{region 'Documentation'}
(*!
<summary>Evaluates captured observations after the scenario has finished.</summary>
*)
{endregion}
METHOD PROTECTED ProcessAssertions
VAR_INPUT
    Enable : BOOL; //! Phase permission supplied by the owning Test Case; FALSE does not authorize progression, while observation may continue.
END_VAR
VAR
    Evaluate : BOOL;
END_VAR
Evaluate := Enable AND FPerformed;
FActiveRun(Enable := Evaluate,
    State := State,
    IN := FActiveRunMatches);
FResetBoundary(Enable := Evaluate,
    State := State,
    IN := FResetBoundaryMatches);
FReservationsReleased(Enable := Evaluate,
    State := State,
    IN := FReservationsReleasedMatches);
FErrorPath(Enable := Evaluate,
    State := State,
    IN := FErrorPathMatches);
FNoLifecycleReset(Enable := Evaluate,
    State := State,
    IN := FNoLifecycleResetMatches);
FNewEpoch(Enable := Evaluate,
    State := State,
    IN := FNewEpochMatches);
FFinalization(Enable := Evaluate,
    State := State,
    IN := FFinalizationMatches);
FConfigurationPreserved(Enable := Evaluate,
    State := State,
    IN := FConfigurationPreservedMatches);
IF Evaluate THEN
    FChecked := TRUE;
END_IF;
END_METHOD

{region 'Documentation'}
(*!
<summary>No Preparation phase is needed.</summary>
*)
{endregion}
METHOD PROTECTED ProcessPreparations
VAR_INPUT
    // SA0033: Required override without Preparation work.
    {attribute 'analysis' := '-33'}
    Enable : BOOL; //! Phase permission supplied by the owning Test Case; FALSE does not authorize progression, while observation may continue.
END_VAR
END_METHOD

{region 'Documentation'}
(*!
<summary>Resets observations and schedules a fresh subject initialization.</summary>
*)
{endregion}
METHOD PROTECTED ProcessReset
FPerformed := FALSE;
FChecked := FALSE;
FPhase := SetupPhase;
FSuite := 0;
FChild := 0;
FSecondChild := 0;
FActiveRun.Reset();
FActiveRunMatches := FALSE;
FResetBoundary.Reset();
FResetBoundaryMatches := FALSE;
FReservationsReleased.Reset();
FReservationsReleasedMatches := FALSE;
FErrorPath.Reset();
FErrorPathMatches := FALSE;
FNoLifecycleReset.Reset();
FNoLifecycleResetMatches := FALSE;
FNewEpoch.Reset();
FNewEpochMatches := FALSE;
FFinalization.Reset();
FFinalizationMatches := FALSE;
FConfigurationPreserved.Reset();
FConfigurationPreservedMatches := FALSE;
CompleteReset();
END_METHOD

{region 'Documentation'}
(*!
<summary>Runs the bounded scenario once before Assertion evaluation.</summary>
*)
{endregion}
METHOD PROTECTED ProcessTests
VAR_INPUT
    Enable : BOOL; //! Phase permission supplied by the owning Test Case; FALSE does not authorize progression, while observation may continue.
END_VAR
IF NOT Enable THEN
    RETURN;
END_IF;
IF FChecked THEN
    CompleteTests();
    RETURN;
END_IF;

IF NOT FPerformed THEN
    StateMachine();
END_IF;
END_METHOD

{region 'Documentation'}
(*!
<summary>Advances the real hierarchy once per cycle and separates reset boundary from error completion.</summary>
*)
{endregion}
METHOD PRIVATE StateMachine
VAR
    EmptyControl : ST_RunControl;
    SeedEvent : ST_Event;
    Published : INT;
END_VAR
CASE FPhase OF
    SetupPhase:
        FControl := EmptyControl;
        IF NOT FSubject.Initialize(Buffer := FEvents,
            FifoControl := FFifo,
            Status := FBufferStatus) THEN
            Error(Message := 'Active reset buffer initialization failed.');
            RETURN;
        END_IF;
        FRoot.BindPublisher(Publisher := FSubject);
        IF NOT FRoot.Initialize(Name := 'ActiveReset',
            EventBuffer := FSubject) THEN
            Error(Message := 'Active reset hierarchy initialization failed.');
            RETURN;
        END_IF;
        FSuite := FRoot.GetTestSuite(Index := FRoot.ChildArrayLowerBound);
        FChild := FRoot.GetTestCase(Index := FRoot.TestCaseLowerBound);
        FSecondChild := FRoot.GetTestCase(Index := FRoot.TestCaseLowerBound + 1);
        IF (FSuite = 0) OR (FChild = 0) OR (FSecondChild = 0) THEN
            Error(Message := 'Active reset hierarchy is incomplete.');
            RETURN;
        END_IF;
        FPhase := AwaitIdlePhase;

    AwaitIdlePhase:
        FRoot(ControlData := FControl);
        IF FRoot.HasError THEN
            Error(Message := 'Active reset hierarchy did not establish Idle.');
            RETURN;
        END_IF;
        IF FRoot.IsReady THEN
            FRoot.RequestStart();
            FPhase := AwaitActivePhase;
        END_IF;

    AwaitActivePhase:
        FRoot(ControlData := FControl);
        IF FRoot.HasError OR FRoot.IsComplete THEN
            Error(Message := 'Hierarchy ended before the active reset precondition.');
            RETURN;
        END_IF;
        IF FChild.State = E_State.Running THEN
            FActiveRunMatches := (FRoot.State = E_State.Running) AND (FSuite.State = E_State.Running)
                AND (FSuite.ReservedEntryCount > 0) AND (FChild.ReservedEntryCount > 0)
                AND (FSubject.ReservedEntryCount > 0);
            SeedEvent := CreateFrameworkEvent(Name := 'ActiveReset',
                ResourceName := 'ActiveResetFixture',
                State := E_State.Running,
                Severity := E_EventSeverity.Info,
                Message := OldEpochMarker);
            Published := FSubject.PublishEvent(Event := SeedEvent);
            FActiveRunMatches := FActiveRunMatches AND (Published > 0);
            FSubject.Arm(Root := FRoot,
                Suite := FSuite,
                Child := FChild);
            FPhase := ResetPhase;
        END_IF;

    ResetPhase:
        FControl.BufferCmd.Reset := TRUE;
        FRoot(ControlData := FControl);
        FResetBoundaryMatches := FSubject.Observed AND FSubject.LifecycleUnchanged
            AND FSubject.EpochCleared AND NOT FControl.BufferCmd.Reset
            AND (FControl.BufferCmd.DeleteSequenceId = 0);
        FReservationsReleasedMatches := FSubject.OwnersReleased
            AND (FSuite.ReservedEntryCount = 0) AND (FChild.ReservedEntryCount = 0)
            AND (FSecondChild.ReservedEntryCount = 0);
        FPhase := AwaitCompletionPhase;

    AwaitCompletionPhase:
        FRoot(ControlData := FControl);
        IF FRoot.IsComplete THEN
            CheckNewEpoch();
            FFinalizationMatches := FFinalizationMatches AND (FRoot.Result = E_Result.Error)
                AND FRoot.HasError;
            FConfigurationPreservedMatches := FRoot.ConfigurationUnchanged AND FRoot.ChildCallsMatch;
            FPerformed := TRUE;
        END_IF;

    ELSE
        Error(Message := 'Unknown active buffer reset phase.');
END_CASE;
END_METHOD

END_FUNCTION_BLOCK

// ---- SelfTests/TestCases/TestSuite_EventBufferReset/Helper/ActiveResetBufferProbe.TcPOU
{region 'Documentation'}
(*!
<summary>Records the synchronous hard-reset boundary before the owner resumes lifecycle processing.</summary>
<description>
Arm captures the real active hierarchy. Reset delegates storage handling unchanged to EventBuffer,
then records cleared metadata and unchanged lifecycle states. Subsequent owner processing may
legitimately publish errors and request Abort; those actions are outside this observation boundary.
Initialization resets are ignored until Arm. The test keeps all referenced objects alive.
</description>
*)
{endregion}
FUNCTION_BLOCK ActiveResetBufferProbe EXTENDS EventBuffer
VAR
    FArmed : BOOL;
    FRoot : REFERENCE TO RunControlIntegrationSubject;
    FSuite : I_TestSuite;
    FChild : I_TestCase;
    FRootState : E_State;
    FSuiteState : E_State;
    FChildState : E_State;
    FLifecycleUnchanged : BOOL;
    FEpochCleared : BOOL;
    FOwnersReleased : BOOL;
    FObserved : BOOL;
END_VAR

{region 'Documentation'}
(*!
<summary>Captures the active hierarchy immediately before the external Buffer Reset.</summary>
*)
{endregion}
METHOD PUBLIC Arm
VAR_INPUT
    Suite : I_TestSuite; //! Borrowed Suite observed across the Reset boundary; keep it alive while armed.
    Child : I_TestCase; //! Borrowed child observed across the Reset boundary; keep it alive while armed.
END_VAR
VAR_IN_OUT
    // SA0167: Borrowed real owner, retained only for state observations.
    {attribute 'analysis' := '-167'}
    Root : RunControlIntegrationSubject; //! Borrowed real Run-Control owner retained for state observations; keep it alive while armed.
END_VAR
FRoot REF= Root;
FSuite := Suite;
FChild := Child;
FRootState := Root.State;
FSuiteState := Suite.State;
FChildState := Child.State;
FLifecycleUnchanged := FALSE;
FEpochCleared := FALSE;
FOwnersReleased := FALSE;
FObserved := FALSE;
FArmed := TRUE;
END_METHOD

{region 'Documentation'}
(*!
<summary>Recorded EpochCleared for command-order verification.</summary>
*)
{endregion}
{attribute 'monitoring' := 'call'}
PROPERTY PUBLIC EpochCleared : BOOL //! Recorded EpochCleared for command-order verification.
GET
EpochCleared := FEpochCleared;
END_GET
END_PROPERTY

{region 'Documentation'}
(*!
<summary>Recorded LifecycleUnchanged for command-order verification.</summary>
*)
{endregion}
{attribute 'monitoring' := 'call'}
PROPERTY PUBLIC LifecycleUnchanged : BOOL //! Recorded LifecycleUnchanged for command-order verification.
GET
LifecycleUnchanged := FLifecycleUnchanged;
END_GET
END_PROPERTY

{region 'Documentation'}
(*!
<summary>Recorded Observed for command-order verification.</summary>
*)
{endregion}
{attribute 'monitoring' := 'call'}
PROPERTY PUBLIC Observed : BOOL //! Recorded Observed for command-order verification.
GET
Observed := FObserved;
END_GET
END_PROPERTY

{region 'Documentation'}
(*!
<summary>Recorded OwnersReleased for command-order verification.</summary>
*)
{endregion}
{attribute 'monitoring' := 'call'}
PROPERTY PUBLIC OwnersReleased : BOOL //! Recorded OwnersReleased for command-order verification.
GET
OwnersReleased := FOwnersReleased;
END_GET
END_PROPERTY

{region 'Documentation'}
(*!
<summary>Delegates real reset and snapshots its immediate effects, not later owner processing.</summary>
*)
{endregion}
METHOD PUBLIC Reset
VAR
    Epoch : ST_EventBufferStatus;
    CurrentFifoStatus : ST_FifoStatus;
END_VAR
IF FArmed THEN
    FOwnersReleased := (FSuite.ReservedEntryCount = 0) AND (FChild.ReservedEntryCount = 0)
        AND (ReservedEntryCount = 0);
END_IF;
SUPER^.Reset();
IF FArmed THEN
    Epoch := Status;
    CurrentFifoStatus := FifoStatus;
    FEpochCleared := CurrentFifoStatus.BufferEmpty AND (CurrentFifoStatus.ElementCount = 0)
        AND (Epoch.SequenceId = 0) AND (Epoch.DeletedSequenceId = 0)
        AND (Epoch.LostEventCount = 0) AND (ReservedEntryCount = 0);
    FLifecycleUnchanged := (FRoot.State = FRootState) AND (FSuite.State = FSuiteState)
        AND (FChild.State = FChildState);
    FObserved := TRUE;
    FArmed := FALSE;
END_IF;
END_METHOD

END_FUNCTION_BLOCK

// ---- SelfTests/TestSuites/TestSuite_AssertionLifecycle.TcPOU
{region 'Documentation'}
(*!
<summary>Checks shared Assertion identity, activity, reset and result-event behavior.</summary>
*)
{endregion}
FUNCTION_BLOCK TestSuite_AssertionLifecycle EXTENDS TestSuiteBase
VAR
    FInitialization : Test_AssertionInitialization;
    FActivity : Test_AssertionActivity;
    FUninitialized : Test_AssertionUninitialized;
    FResetReuse : Test_AssertionResetReuse;
    FEscalation : Test_AssertionEscalation;
    FTestCases : ARRAY[1..TestCaseCapacity] OF I_TestCase;
END_VAR
VAR CONSTANT
    TestCaseCapacity : UINT := 5;
END_VAR

SUPER^();

{region 'Documentation'}
(*!
<summary>Initializes and registers the five isolated Assertion lifecycle scenarios.</summary>
*)
{endregion}
METHOD PROTECTED Configure
VAR_IN_OUT
    // SA0167: Borrowed owner builder; no temporary instance is created.
    {attribute 'analysis' := '-167'}
    Builder : TestSuiteConfigurationBuilder; //! Borrowed owner configuration builder used only during this Configure call; register this owner's concrete children.
END_VAR
VAR
    TestConfig : ST_TestCaseConfig;
END_VAR
Builder.Initialize(Mode := E_OrchestrationMode.Serial,
    TestCases := FTestCases);
FInitialization.Initialize(Parent := THIS^,
    TestName := 'Initialization',
    Config := TestConfig);
Builder.Register(TestCase := FInitialization);
FActivity.Initialize(Parent := THIS^,
    TestName := 'Activity',
    Config := TestConfig);
Builder.Register(TestCase := FActivity);
FUninitialized.Initialize(Parent := THIS^,
    TestName := 'Uninitialized',
    Config := TestConfig);
Builder.Register(TestCase := FUninitialized);
FResetReuse.Initialize(Parent := THIS^,
    TestName := 'ResetReuse',
    Config := TestConfig);
Builder.Register(TestCase := FResetReuse);
FEscalation.Initialize(Parent := THIS^,
    TestName := 'Escalation',
    Config := TestConfig);
Builder.Register(TestCase := FEscalation);
END_METHOD

{region 'Documentation'}
(*!
<summary>Returns a registered scenario using its original array index.</summary>
*)
{endregion}
METHOD PUBLIC GetTestCase : I_TestCase //! Typed child interface at the original array index; zero when no entry is available.
VAR_INPUT
    Index : DINT; //! Original occupied child-array index, rather than an ordinal position.
END_VAR
GetTestCase := 0;
IF (ChildCount = 0) OR (Index < ChildArrayLowerBound)
    OR (DINT_TO_LINT(Index) >= DINT_TO_LINT(ChildArrayLowerBound) + UINT_TO_LINT(ChildCount)) THEN
    RETURN;
END_IF;
GetTestCase := FTestCases[Index];
END_METHOD

{region 'Documentation'}
(*!
<summary>Calls each owned scenario once per initialized Suite cycle.</summary>
*)
{endregion}
METHOD PROTECTED ProcessTestCases
FInitialization();
FActivity();
FUninitialized();
FResetReuse();
FEscalation();
END_METHOD

END_FUNCTION_BLOCK

// ---- SelfTests/TestCases/TestSuite_AssertionLifecycle/Test_AssertionInitialization.TcPOU
{region 'Documentation'}
(*!
<summary>Checks Assertion identity validation and deferred reset dispatch.</summary>
<description>
Each attempt changes one identity/configuration condition. Initialize is checked before
any FB call; three later calls verify reset dispatch, valid activity or rejected passivity.
Checking Assertions latch every attempt, while intentional diagnostics stay local.
Publisher checks cover zero rejection, explicit replacement and unchanged lifecycle/history
before and after subject calls. A separate untouched Assertion verifies the lazy default.
Repeated runs use the same subject and reinitialize it; they do not claim fresh memory.
</description>
*)
{endregion}
FUNCTION_BLOCK Test_AssertionInitialization EXTENDS TestCaseBase
VAR
    FSubject : AssertionLifecycleSubject;
    FDefaultSubject : AssertTrue;
    FAlternativeCapture : EventBuffer;
    FAlternativeEvents : ARRAY[1..CaptureLength] OF ST_Event;
    FAlternativeFifo : ST_FifoStatus;
    FAlternativeStatus : ST_EventBufferStatus;
    FParent : AssertionParentIdentity;
    FCapture : EventBuffer;
    FEvents : ARRAY[1..CaptureLength] OF ST_Event;
    FCaptureFifo : ST_FifoStatus;
    FCaptureStatus : ST_EventBufferStatus;
    FAttempt : UINT;
    FCall : UINT;
    FAttemptStarted : BOOL;
    FExpectedInitialized : BOOL;
    FExpectedObserveFirstCycle : BOOL;
    FExpectedName : STRING(GVL_Constants.NameLength);
    FExpectedResource : STRING(GVL_Constants.ResourceNameLength);
    FExpectedEvents : UDINT;
    FObservationReady : BOOL;
    FChecked : BOOL;
END_VAR
VAR
    FPublisherBinding : AssertTrue;
    FPublisherBindingMatches : BOOL;
    FInitialization : AssertTrue;
    FInitializationMatches : BOOL;
    FIdentity : AssertTrue;
    FIdentityMatches : BOOL;
    FSettings : AssertTrue;
    FSettingsMatches : BOOL;
    FDispatch : AssertTrue;
    FDispatchMatches : BOOL;
    FActivity : AssertTrue;
    FActivityMatches : BOOL;
    FDiagnostics : AssertTrue;
    FDiagnosticsMatches : BOOL;
    FCaptureIntegrity : AssertTrue;
    FCaptureIntegrityMatches : BOOL;
END_VAR
VAR CONSTANT
    CaptureLength : UINT := 8;
    DefaultSettings : UINT := 1;
    DottedSuffix : UINT := 2;
    ExactCapacity : UINT := 3;
    OverCapacity : UINT := 4;
    MissingParent : UINT := 5;
    EmptySuffix : UINT := 6;
    InvalidParent : UINT := 7;
    NonAsciiSuffix : UINT := 8;
    ExplicitSettings : UINT := 9;
    LastAttempt : UINT := ExplicitSettings;
    ResetCall : UINT := 1;
    SecondCheckCall : UINT := 3;
    ResetSampleValue : UINT := 17;
END_VAR

SUPER^();

{region 'Documentation'}
(*!
<summary>Collects only outer checking Assertions, never intentional subject findings.</summary>
*)
{endregion}
METHOD PROTECTED AggregateResults
VAR_INPUT
    Aggregator : I_ResultAggregator; //! Borrowed result sink owned by the outer Test Case; add this test's checking Assertions without resetting or retaining the sink.
END_VAR
Aggregator.AddProvider(Provider := FPublisherBinding);
Aggregator.AddProvider(Provider := FInitialization);
Aggregator.AddProvider(Provider := FIdentity);
Aggregator.AddProvider(Provider := FSettings);
Aggregator.AddProvider(Provider := FDispatch);
Aggregator.AddProvider(Provider := FActivity);
Aggregator.AddProvider(Provider := FDiagnostics);
Aggregator.AddProvider(Provider := FCaptureIntegrity);
END_METHOD

{region 'Documentation'}
(*!
<summary>Varies one setup condition and observes Initialize before cyclic processing.</summary>
*)
{endregion}
METHOD PRIVATE BeginAttempt
VAR
    Parent : I_TestCase;
    ParentName : STRING(GVL_Constants.NameLength);
    LocalName : STRING(GVL_Constants.NameLength);
    FullName : STRING(2 * GVL_Constants.NameLength + 1);
    Initialized : BOOL;
    SuffixLength : INT;
    Index : INT;
END_VAR
IF NOT FCapture.Initialize(Buffer := FEvents,
    FifoControl := FCaptureFifo,
    Status := FCaptureStatus) THEN
    Error(Message := 'Assertion initialization capture setup failed.');
    RETURN;
END_IF;

IF NOT FAlternativeCapture.Initialize(Buffer := FAlternativeEvents,
    FifoControl := FAlternativeFifo,
    Status := FAlternativeStatus) THEN
    Error(Message := 'Alternative Assertion publisher setup failed.');
    RETURN;
END_IF;

CheckPublisherBinding();
ParentName := 'Root.Suite.Case';
LocalName := 'Subject';
FExpectedInitialized := TRUE;
FExpectedObserveFirstCycle := TRUE;
FExpectedResource := '';
CASE FAttempt OF
    DefaultSettings:
        LocalName := 'Subject';
    DottedSuffix:
        LocalName := 'Value.With.Detail';
    ExactCapacity, OverCapacity:
        LocalName := '';
        SuffixLength := UINT_TO_INT(GVL_Constants.NameLength) - LEN(ParentName) - 1;
        IF FAttempt = OverCapacity THEN
            SuffixLength := SuffixLength + 1;
            FExpectedInitialized := FALSE;
        END_IF;
        FOR Index := 1 TO SuffixLength DO
            LocalName := CONCAT(LocalName, 'x');
        END_FOR;
    MissingParent:
        FExpectedInitialized := FALSE;
    EmptySuffix:
        LocalName := '';
        FExpectedInitialized := FALSE;
    InvalidParent:
        ParentName := 'Root..Case';
        FExpectedInitialized := FALSE;
    NonAsciiSuffix:
        // SA0175: Deliberately invalid non-ASCII identity input for the rejection test.
        {analysis -175}
        LocalName := '$E4';
        {analysis +175}
        FExpectedInitialized := FALSE;
    ExplicitSettings:
        FExpectedResource := 'Resource';
        FExpectedObserveFirstCycle := FALSE;
ELSE
    Error(Message := 'Unknown Assertion initialization attempt.');
    RETURN;
END_CASE;

FParent.SetIdentity(Value := ParentName);
Parent := FParent;
IF FAttempt = MissingParent THEN
    Parent := 0;
    FExpectedName := LocalName;
ELSE
    FullName := CONCAT(CONCAT(ParentName, '.'), LocalName);
    // SA0175: The expected diagnostic projection is deliberately bounded ASCII-byte truncation.
    {analysis -175}
    FExpectedName := LEFT(FullName, UINT_TO_INT(GVL_Constants.NameLength));
    {analysis +175}
END_IF;

FSubject.ClearTrace();
IF FAttempt = ExplicitSettings THEN
    Initialized := FSubject.Initialize(Parent := Parent,
        AssertionName := LocalName,
        ResourceName := FExpectedResource,
        ObserveFirstCycle := FExpectedObserveFirstCycle);
ELSE
    Initialized := FSubject.Initialize(Parent := Parent,
        AssertionName := LocalName);
END_IF;
FInitializationMatches := (Initialized = FExpectedInitialized)
    AND (FSubject.IsInitialized = FExpectedInitialized)
    AND (FSubject.Result = E_Result.NotEvaluated);
FIdentityMatches := TRUE;
FSettingsMatches := TRUE;
IF FAttempt <> MissingParent THEN
    FIdentityMatches := FSubject.Name = FExpectedName;
    FSettingsMatches := (FSubject.ResourceName = FExpectedResource)
        AND (FSubject.ObserveFirstCycle = FExpectedObserveFirstCycle);
END_IF;
FDispatchMatches := (FSubject.ResetCallCount = 0) AND (FSubject.AssertCallCount = 0);
FActivityMatches := NOT FSubject.Enabled
    AND NOT FSubject.ObservationActive AND NOT FSubject.EvaluationActive;
FExpectedEvents := 0;
FDiagnosticsMatches := TRUE;
IF NOT FExpectedInitialized THEN
    FExpectedEvents := 1;
    FDiagnosticsMatches := (FEvents[1].Name = FExpectedName)
        AND (FEvents[1].OwnerScope = E_OwnerScope.Framework)
        AND (FEvents[1].EventType = E_EventType.Framework)
        AND (FEvents[1].Severity = E_EventSeverity.Error)
        AND (FEvents[1].State = E_State.Uninitialized);
END_IF;
FDiagnosticsMatches := FDiagnosticsMatches AND (FCaptureStatus.SequenceId = FExpectedEvents);
FCaptureIntegrityMatches := FCaptureStatus.LostEventCount = 0;
FAttemptStarted := TRUE;
FCall := ResetCall;
END_METHOD

{region 'Documentation'}
(*!
<summary>Checks binding without changing subject lifecycle, history or event counts.</summary>
*)
{endregion}
METHOD PRIVATE CheckPublisherBinding
VAR
    PrimaryPublisher : I_EventPublisher;
    AlternativePublisher : I_EventPublisher;
    DefaultPublisher : I_EventPublisher;
    ResultBefore : E_Result;
    InitializedBefore : BOOL;
    EnabledBefore : BOOL;
    ObservationBefore : BOOL;
    EvaluationBefore : BOOL;
    NameBefore : STRING(GVL_Constants.NameLength);
    SequenceBefore : UDINT;
    AlternativeSequenceBefore : UDINT;
END_VAR
PrimaryPublisher := FCapture;
AlternativePublisher := FAlternativeCapture;
DefaultPublisher := GVL_EventBuffer.Publisher;
FDefaultSubject.BindPublisher(Publisher := 0);
FPublisherBindingMatches := FPublisherBindingMatches
    AND (FDefaultSubject.EventPublisher = DefaultPublisher);

ResultBefore := FSubject.Result;
InitializedBefore := FSubject.IsInitialized;
EnabledBefore := FSubject.Enabled;
ObservationBefore := FSubject.ObservationActive;
EvaluationBefore := FSubject.EvaluationActive;
NameBefore := FSubject.Name;
SequenceBefore := FCaptureStatus.SequenceId;
AlternativeSequenceBefore := FAlternativeStatus.SequenceId;

FSubject.BindPublisher(Publisher := AlternativePublisher);
FPublisherBindingMatches := FPublisherBindingMatches
    AND (FSubject.EventPublisher = AlternativePublisher);
FSubject.BindPublisher(Publisher := 0);
FPublisherBindingMatches := FPublisherBindingMatches
    AND (FSubject.EventPublisher = AlternativePublisher);
FSubject.BindPublisher(Publisher := PrimaryPublisher);
FPublisherBindingMatches := FPublisherBindingMatches
    AND (FSubject.EventPublisher = PrimaryPublisher)
    AND (FSubject.Result = ResultBefore)
    AND (FSubject.IsInitialized = InitializedBefore)
    AND (FSubject.Enabled = EnabledBefore)
    AND (FSubject.ObservationActive = ObservationBefore)
    AND (FSubject.EvaluationActive = EvaluationBefore)
    AND (FSubject.Name = NameBefore)
    AND (FCaptureStatus.SequenceId = SequenceBefore)
    AND (FAlternativeStatus.SequenceId = AlternativeSequenceBefore);
END_METHOD

{region 'Documentation'}
(*!
<summary>Configures checking Assertions; subject actions remain in the test script.</summary>
*)
{endregion}
METHOD PROTECTED Configure
FPreparationStateCount := 0;
FTestStateCount := 1;
FPublisherBinding.Initialize(Parent := THIS^,
    AssertionName := 'PublisherBinding');
FInitialization.Initialize(Parent := THIS^,
    AssertionName := 'Initialization');
FIdentity.Initialize(Parent := THIS^,
    AssertionName := 'Identity');
FSettings.Initialize(Parent := THIS^,
    AssertionName := 'Settings');
FDispatch.Initialize(Parent := THIS^,
    AssertionName := 'Dispatch');
FActivity.Initialize(Parent := THIS^,
    AssertionName := 'Activity');
FDiagnostics.Initialize(Parent := THIS^,
    AssertionName := 'Diagnostics');
FCaptureIntegrity.Initialize(Parent := THIS^,
    AssertionName := 'CaptureIntegrity');
FSubject.BindPublisher(Publisher := FCapture);
END_METHOD

{region 'Documentation'}
(*!
<summary>Checks reset and subsequent dispatch using one subject call per cycle.</summary>
*)
{endregion}
METHOD PRIVATE ObserveCall
VAR
    ExpectedActive : BOOL;
END_VAR
FSubject(Enable := TRUE,
    State := E_State.Running,
    Sample := ResetSampleValue);
FDispatchMatches := FDispatchMatches
    AND (FSubject.ResetCallCount = 1) AND (FSubject.ResetSample = ResetSampleValue);
IF FCall = ResetCall THEN
    FDispatchMatches := FDispatchMatches AND (FSubject.AssertCallCount = 0)
        AND (FSubject.ObservedSample = 0);
    FActivityMatches := FActivityMatches AND FSubject.Enabled
        AND NOT FSubject.ObservationActive AND NOT FSubject.EvaluationActive
        AND (FSubject.Result = E_Result.NotEvaluated);
ELSIF FExpectedInitialized THEN
    FDispatchMatches := FDispatchMatches AND (FSubject.AssertCallCount = FCall - 1);
    ExpectedActive := FExpectedObserveFirstCycle OR (FCall = SecondCheckCall);
    FActivityMatches := FActivityMatches AND FSubject.Enabled
        AND (FSubject.ObservationActive = ExpectedActive)
        AND (FSubject.EvaluationActive = ExpectedActive);
    IF ExpectedActive THEN
        FActivityMatches := FActivityMatches AND (FSubject.Result = E_Result.Passed);
    ELSE
        FActivityMatches := FActivityMatches AND (FSubject.Result = E_Result.NotEvaluated);
    END_IF;
ELSE
    FDispatchMatches := FDispatchMatches AND (FSubject.AssertCallCount = 0);
    FActivityMatches := FActivityMatches AND NOT FSubject.ObservationActive
        AND NOT FSubject.EvaluationActive AND (FSubject.Result = E_Result.NotEvaluated);
END_IF;
FDiagnosticsMatches := FDiagnosticsMatches AND (FCaptureStatus.SequenceId = FExpectedEvents);
FCaptureIntegrityMatches := FCaptureIntegrityMatches AND (FCaptureStatus.LostEventCount = 0);
CheckPublisherBinding();
FObservationReady := TRUE;
END_METHOD

{region 'Documentation'}
(*!
<summary>Completes abort without asynchronous resources.</summary>
*)
{endregion}
METHOD PROTECTED ProcessAbort
VAR_INPUT
    Enable : BOOL; //! Phase permission supplied by the owning Test Case; FALSE does not authorize progression, while observation may continue.
END_VAR
IF Enable THEN
    CompleteAbort();
END_IF;
END_METHOD

{region 'Documentation'}
(*!
<summary>Latches checked observations before the next script step may proceed.</summary>
*)
{endregion}
METHOD PROTECTED ProcessAssertions
VAR_INPUT
    Enable : BOOL; //! Phase permission supplied by the owning Test Case; FALSE does not authorize progression, while observation may continue.
END_VAR
VAR
    Evaluate : BOOL;
END_VAR
Evaluate := Enable AND FObservationReady;
FPublisherBinding(Enable := Evaluate,
    State := State,
    IN := FPublisherBindingMatches);
FInitialization(Enable := Evaluate,
    State := State,
    IN := FInitializationMatches);
FIdentity(Enable := Evaluate,
    State := State,
    IN := FIdentityMatches);
FSettings(Enable := Evaluate,
    State := State,
    IN := FSettingsMatches);
FDispatch(Enable := Evaluate,
    State := State,
    IN := FDispatchMatches);
FActivity(Enable := Evaluate,
    State := State,
    IN := FActivityMatches);
FDiagnostics(Enable := Evaluate,
    State := State,
    IN := FDiagnosticsMatches);
FCaptureIntegrity(Enable := Evaluate,
    State := State,
    IN := FCaptureIntegrityMatches);
IF Evaluate THEN
    FChecked := TRUE;
END_IF;
END_METHOD

{region 'Documentation'}
(*!
<summary>No Preparation phase is required.</summary>
*)
{endregion}
METHOD PROTECTED ProcessPreparations
VAR_INPUT
    // SA0033: Required hook; this test has no Preparation phase.
    {attribute 'analysis' := '-33'}
    Enable : BOOL; //! Phase permission supplied by the owning Test Case; FALSE does not authorize progression, while observation may continue.
END_VAR
END_METHOD

{region 'Documentation'}
(*!
<summary>Restarts the script and resets the checking Assertions.</summary>
*)
{endregion}
METHOD PROTECTED ProcessReset
FPublisherBinding.Reset();
FPublisherBindingMatches := TRUE;
FAttempt := DefaultSettings;
FCall := ResetCall;
FAttemptStarted := FALSE;
FObservationReady := FALSE;
FChecked := FALSE;
FInitialization.Reset();
FInitializationMatches := TRUE;
FIdentity.Reset();
FIdentityMatches := TRUE;
FSettings.Reset();
FSettingsMatches := TRUE;
FDispatch.Reset();
FDispatchMatches := TRUE;
FActivity.Reset();
FActivityMatches := TRUE;
FDiagnostics.Reset();
FDiagnosticsMatches := TRUE;
FCaptureIntegrity.Reset();
FCaptureIntegrityMatches := TRUE;
CompleteReset();
END_METHOD

{region 'Documentation'}
(*!
<summary>Advances one bounded script step per active PLC cycle.</summary>
*)
{endregion}
METHOD PROTECTED ProcessTests
VAR_INPUT
    Enable : BOOL; //! Phase permission supplied by the owning Test Case; FALSE does not authorize progression, while observation may continue.
END_VAR
IF NOT Enable THEN
    RETURN;
END_IF;
IF FChecked THEN
    FChecked := FALSE;
    FObservationReady := FALSE;
    IF FCall = SecondCheckCall THEN
        IF FAttempt = LastAttempt THEN
            CompleteTests();
            RETURN;
        END_IF;
        FAttempt := FAttempt + 1;
        FAttemptStarted := FALSE;
    ELSE
        FCall := FCall + 1;
    END_IF;
END_IF;
IF NOT FAttemptStarted THEN
    BeginAttempt();
    RETURN;
END_IF;
ObserveCall();
END_METHOD

END_FUNCTION_BLOCK

// ---- SelfTests/TestCases/TestSuite_AssertionLifecycle/Helper/AssertionLifecycleSubject.TcPOU
{region 'Documentation'}
(*!
<summary>Exposes calls and activity gates of AssertionBase without replacing its processing.</summary>
<description>
Bind the local publisher before Initialize. The inherited body owns initialization,
reset priority and activity history. Assert records both gates and a bounded sample;
active evaluation dispatches the selected inherited finding method without a result guard.
This deliberately exercises base-owned suppression. Counters are cumulative until ClearTrace.
ResetAssertion clears the sample and records the input available on the reset call.
The outer test owns expectations; this subject does not compute expected gates.
</description>
*)
{endregion}
FUNCTION_BLOCK AssertionLifecycleSubject EXTENDS AssertionBase
VAR_INPUT
    Sample : UINT := 0; //! Controlled sample captured only while observation is active.
    Finding : E_Result := E_Result.Passed; //! Passed, Failed or Error finding dispatched only while evaluation is active.
    FindingMessage : STRING(GVL_Constants.MessageLength) := 'Controlled finding.'; //! Diagnostic text supplied to the selected Fail or Error operation.
END_VAR
VAR_OUTPUT
    AssertCallCount : UINT; //! Cumulative Assert-hook invocations since ClearTrace.
    ResetCallCount : UINT; //! Cumulative ResetAssertion-hook invocations since ClearTrace.
    ObservationCount : UINT; //! Cumulative Assert calls with the observation gate active since ClearTrace.
    EvaluationCount : UINT; //! Cumulative Assert calls with the evaluation gate active since ClearTrace.
    ObservedSample : UINT; //! Last Sample accepted while observation was active; ResetAssertion clears it.
    ResetSample : UINT; //! Sample present at the latest ResetAssertion call.
    ObservationDuringAssert : BOOL; //! Observation gate recorded on the latest Assert-hook entry.
    EvaluationDuringAssert : BOOL; //! Evaluation gate recorded on the latest Assert-hook entry.
END_VAR

SUPER^();

{region 'Documentation'}
(*!
<summary>Records inherited gates and evaluates only when permitted.</summary>
*)
{endregion}
METHOD PROTECTED Assert
AssertCallCount := AssertCallCount + 1;
ObservationDuringAssert := ObservationActive;
EvaluationDuringAssert := EvaluationActive;
IF ObservationDuringAssert THEN
    ObservationCount := ObservationCount + 1;
    ObservedSample := Sample;
END_IF;
IF EvaluationDuringAssert THEN
    EvaluationCount := EvaluationCount + 1;
    CASE Finding OF
        E_Result.Passed:
            Pass();
        E_Result.Failed:
            Fail(Message := FindingMessage);
        E_Result.Error:
            Error(Message := FindingMessage);
    ELSE
        RETURN;
    END_CASE;
END_IF;
END_METHOD

{region 'Documentation'}
(*!
<summary>Clears only test instrumentation; never changes inherited Assertion state.</summary>
*)
{endregion}
METHOD PUBLIC ClearTrace
AssertCallCount := 0;
ResetCallCount := 0;
ObservationCount := 0;
EvaluationCount := 0;
ObservedSample := 0;
ResetSample := 0;
ObservationDuringAssert := FALSE;
EvaluationDuringAssert := FALSE;
END_METHOD

{region 'Documentation'}
(*!
<summary>Records one reset with bound inputs and clears the observation sample.</summary>
*)
{endregion}
METHOD PROTECTED ResetAssertion
ResetCallCount := ResetCallCount + 1;
ResetSample := Sample;
ObservedSample := 0;
END_METHOD

END_FUNCTION_BLOCK

// ---- SelfTests/TestCases/TestSuite_AssertionLifecycle/Helper/AssertionParentIdentity.TcPOU
{region 'Documentation'}
(*!
<summary>Supplies controlled parent identity for Assertion initialization tests.</summary>
<description>
Only Name is consumed by the subject. SetIdentity deliberately admits malformed names
to exercise the subject boundary. This local mock is never scheduled as a Test Case.
</description>
*)
{endregion}
FUNCTION_BLOCK AssertionParentIdentity EXTENDS TestCaseMock

SUPER^();

{region 'Documentation'}
(*!
<summary>Sets the parent name before the subject reads it; no lifecycle work.</summary>
*)
{endregion}
METHOD PUBLIC SetIdentity
VAR_INPUT
    Value : STRING(GVL_Constants.NameLength); //! Identity-only parent name retained for isolated Assertion initialization.
END_VAR
FName := Value;
END_METHOD

END_FUNCTION_BLOCK

// ---- SelfTests/TestCases/TestSuite_AssertionLifecycle/Test_AssertionActivity.TcPOU
{region 'Documentation'}
(*!
<summary>Checks both Assertion activity strategies with literal cycle expectations.</summary>
<description>
The Suite selects ObserveFirstCycle before initialization and keeps it fixed.
Each active cycle calls each subject once. The script includes independent Evaluate
while disabled and on the first excluded observation call, plus disable/re-enable.
Expected steps are specified here, not obtained from the subject's gate formulas.
Initial reset consumes bound inputs and suppresses both gates even when requested.
</description>
*)
{endregion}
FUNCTION_BLOCK Test_AssertionActivity EXTENDS TestCaseBase
VAR_INPUT
    ObserveFirstCycle : BOOL := TRUE; //! First-cycle observation strategy selected before initialization and held fixed by the containing Suite.
END_VAR
VAR
    FDirect : AssertionLifecycleSubject;
    FExplicit : AssertionEvaluationSubject;
    FCapture : EventBuffer;
    FEvents : ARRAY[1..CaptureLength] OF ST_Event;
    FCaptureFifo : ST_FifoStatus;
    FCaptureStatus : ST_EventBufferStatus;
    FStep : UINT;
    FObservationReady : BOOL;
    FChecked : BOOL;
    FEnable : BOOL;
    FEvaluate : BOOL;
    FExpectedObservation : BOOL;
    FExpectedExplicitEvaluation : BOOL;
    FExpectedObservationCount : UINT;
    FExpectedExplicitCount : UINT;
END_VAR
VAR
    FInitialization : AssertTrue;
    FInitializationMatches : BOOL;
    FEnabled : AssertTrue;
    FEnabledMatches : BOOL;
    FObservation : AssertTrue;
    FObservationMatches : BOOL;
    FDirectEvaluation : AssertTrue;
    FDirectEvaluationMatches : BOOL;
    FExplicitEvaluation : AssertTrue;
    FExplicitEvaluationMatches : BOOL;
    FHookDispatch : AssertTrue;
    FHookDispatchMatches : BOOL;
    FStableProperties : AssertTrue;
    FStablePropertiesMatches : BOOL;
    FNoFindings : AssertTrue;
    FNoFindingsMatches : BOOL;
END_VAR
VAR CONSTANT
    CaptureLength : UINT := 8;
    InitializeSubjects : UINT := 0;
    ConsumeInitialReset : UINT := 1;
    DisabledCall : UINT := 2;
    FirstEnabledCall : UINT := 3;
    ObservationOnly : UINT := 4;
    EvaluationOnly : UINT := 5;
    FirstReenabledCall : UINT := 6;
    ContinuedCall : UINT := 7;
END_VAR

SUPER^();

{region 'Documentation'}
(*!
<summary>Collects only outer checking Assertions, never intentional subject findings.</summary>
*)
{endregion}
METHOD PROTECTED AggregateResults
VAR_INPUT
    Aggregator : I_ResultAggregator; //! Borrowed result sink owned by the outer Test Case; add this test's checking Assertions without resetting or retaining the sink.
END_VAR
Aggregator.AddProvider(Provider := FInitialization);
Aggregator.AddProvider(Provider := FEnabled);
Aggregator.AddProvider(Provider := FObservation);
Aggregator.AddProvider(Provider := FDirectEvaluation);
Aggregator.AddProvider(Provider := FExplicitEvaluation);
Aggregator.AddProvider(Provider := FHookDispatch);
Aggregator.AddProvider(Provider := FStableProperties);
Aggregator.AddProvider(Provider := FNoFindings);
END_METHOD

{region 'Documentation'}
(*!
<summary>Configures checking Assertions; subject actions remain in the test script.</summary>
*)
{endregion}
METHOD PROTECTED Configure
FPreparationStateCount := 0;
FTestStateCount := 1;
FInitialization.Initialize(Parent := THIS^,
    AssertionName := 'Initialization');
FEnabled.Initialize(Parent := THIS^,
    AssertionName := 'Enabled');
FObservation.Initialize(Parent := THIS^,
    AssertionName := 'Observation');
FDirectEvaluation.Initialize(Parent := THIS^,
    AssertionName := 'DirectEvaluation');
FExplicitEvaluation.Initialize(Parent := THIS^,
    AssertionName := 'ExplicitEvaluation');
FHookDispatch.Initialize(Parent := THIS^,
    AssertionName := 'HookDispatch');
FStableProperties.Initialize(Parent := THIS^,
    AssertionName := 'StableProperties');
FNoFindings.Initialize(Parent := THIS^,
    AssertionName := 'NoFindings');
FDirect.BindPublisher(Publisher := FCapture);
FExplicit.BindPublisher(Publisher := FCapture);
END_METHOD

{region 'Documentation'}
(*!
<summary>Initializes both subjects and checks their immediately inactive state.</summary>
*)
{endregion}
METHOD PRIVATE InitializeActivitySubjects
VAR
    DirectInitialized : BOOL;
    ExplicitInitialized : BOOL;
END_VAR
IF NOT FCapture.Initialize(Buffer := FEvents,
    FifoControl := FCaptureFifo,
    Status := FCaptureStatus) THEN
    Error(Message := 'Assertion activity capture setup failed.');
    RETURN;
END_IF;
FDirect.ClearTrace();
FExplicit.ClearTrace();
DirectInitialized := FDirect.Initialize(Parent := THIS^,
    AssertionName := 'DirectSubject',
    ObserveFirstCycle := ObserveFirstCycle);
ExplicitInitialized := FExplicit.Initialize(Parent := THIS^,
    AssertionName := 'ExplicitSubject',
    ObserveFirstCycle := ObserveFirstCycle);
FInitializationMatches := DirectInitialized AND ExplicitInitialized
    AND FDirect.IsInitialized AND FExplicit.IsInitialized
    AND NOT FDirect.Enabled AND NOT FExplicit.Enabled
    AND NOT FDirect.ObservationActive AND NOT FExplicit.ObservationActive
    AND NOT FDirect.EvaluationActive AND NOT FExplicit.EvaluationActive
    AND (FDirect.ResetCallCount = 0) AND (FExplicit.ResetCallCount = 0)
    AND (FDirect.Result = E_Result.NotEvaluated) AND (FExplicit.Result = E_Result.NotEvaluated);
FStep := ConsumeInitialReset;
END_METHOD

{region 'Documentation'}
(*!
<summary>Executes both subjects once and checks gates, hook counts and retained results.</summary>
*)
{endregion}
METHOD PRIVATE ObserveCall
FDirect(Enable := FEnable,
    State := E_State.Running,
    Sample := FStep);
FExplicit(Enable := FEnable,
    Evaluate := FEvaluate,
    State := E_State.Running,
    Sample := FStep);
IF FExpectedObservation THEN
    FExpectedObservationCount := FExpectedObservationCount + 1;
END_IF;
IF FExpectedExplicitEvaluation THEN
    FExpectedExplicitCount := FExpectedExplicitCount + 1;
END_IF;

FEnabledMatches := (FDirect.Enabled = FEnable) AND (FExplicit.Enabled = FEnable);
FObservationMatches := (FDirect.ObservationActive = FExpectedObservation)
    AND (FExplicit.ObservationActive = FExpectedObservation)
    AND (FDirect.ObservationCount = FExpectedObservationCount)
    AND (FExplicit.ObservationCount = FExpectedObservationCount);
FDirectEvaluationMatches := (FDirect.EvaluationActive = FExpectedObservation)
    AND (FDirect.EvaluationCount = FExpectedObservationCount);
FExplicitEvaluationMatches := (FExplicit.EvaluationActive = FExpectedExplicitEvaluation)
    AND (FExplicit.EvaluationCount = FExpectedExplicitCount);
IF FExpectedObservationCount = 0 THEN
    FDirectEvaluationMatches := FDirectEvaluationMatches AND (FDirect.Result = E_Result.NotEvaluated);
ELSE
    FDirectEvaluationMatches := FDirectEvaluationMatches AND (FDirect.Result = E_Result.Passed);
END_IF;
IF FExpectedExplicitCount = 0 THEN
    FExplicitEvaluationMatches := FExplicitEvaluationMatches AND (FExplicit.Result = E_Result.NotEvaluated);
ELSE
    FExplicitEvaluationMatches := FExplicitEvaluationMatches AND (FExplicit.Result = E_Result.Passed);
END_IF;

FHookDispatchMatches := (FDirect.ResetCallCount = 1) AND (FExplicit.ResetCallCount = 1)
    AND (FDirect.ResetSample = ConsumeInitialReset) AND (FExplicit.ResetSample = ConsumeInitialReset)
    AND (FDirect.AssertCallCount = FStep - ConsumeInitialReset)
    AND (FExplicit.AssertCallCount = FStep - ConsumeInitialReset);
FStablePropertiesMatches := TRUE;
IF FStep <> ConsumeInitialReset THEN
    FStablePropertiesMatches := (FDirect.ObservationDuringAssert = FDirect.ObservationActive)
        AND (FDirect.EvaluationDuringAssert = FDirect.EvaluationActive)
        AND (FExplicit.ObservationDuringAssert = FExplicit.ObservationActive)
        AND (FExplicit.EvaluationDuringAssert = FExplicit.EvaluationActive);
END_IF;
// Repeat reads must neither advance history nor change the last call's effective gates.
FStablePropertiesMatches := FStablePropertiesMatches
    AND (FDirect.ObservationActive = FExpectedObservation)
    AND (FDirect.EvaluationActive = FExpectedObservation)
    AND (FExplicit.ObservationActive = FExpectedObservation)
    AND (FExplicit.EvaluationActive = FExpectedExplicitEvaluation);
FNoFindingsMatches := (FCaptureStatus.SequenceId = 0) AND (FCaptureStatus.LostEventCount = 0);
FObservationReady := TRUE;
END_METHOD

{region 'Documentation'}
(*!
<summary>Completes abort without asynchronous resources.</summary>
*)
{endregion}
METHOD PROTECTED ProcessAbort
VAR_INPUT
    Enable : BOOL; //! Phase permission supplied by the owning Test Case; FALSE does not authorize progression, while observation may continue.
END_VAR
IF Enable THEN
    CompleteAbort();
END_IF;
END_METHOD

{region 'Documentation'}
(*!
<summary>Latches checked observations before the next script step may proceed.</summary>
*)
{endregion}
METHOD PROTECTED ProcessAssertions
VAR_INPUT
    Enable : BOOL; //! Phase permission supplied by the owning Test Case; FALSE does not authorize progression, while observation may continue.
END_VAR
VAR
    Evaluate : BOOL;
END_VAR
Evaluate := Enable AND FObservationReady;
FInitialization(Enable := Evaluate,
    State := State,
    IN := FInitializationMatches);
FEnabled(Enable := Evaluate,
    State := State,
    IN := FEnabledMatches);
FObservation(Enable := Evaluate,
    State := State,
    IN := FObservationMatches);
FDirectEvaluation(Enable := Evaluate,
    State := State,
    IN := FDirectEvaluationMatches);
FExplicitEvaluation(Enable := Evaluate,
    State := State,
    IN := FExplicitEvaluationMatches);
FHookDispatch(Enable := Evaluate,
    State := State,
    IN := FHookDispatchMatches);
FStableProperties(Enable := Evaluate,
    State := State,
    IN := FStablePropertiesMatches);
FNoFindings(Enable := Evaluate,
    State := State,
    IN := FNoFindingsMatches);
IF Evaluate THEN
    FChecked := TRUE;
END_IF;
END_METHOD

{region 'Documentation'}
(*!
<summary>No Preparation phase is required.</summary>
*)
{endregion}
METHOD PROTECTED ProcessPreparations
VAR_INPUT
    // SA0033: Required hook; this test has no Preparation phase.
    {attribute 'analysis' := '-33'}
    Enable : BOOL; //! Phase permission supplied by the owning Test Case; FALSE does not authorize progression, while observation may continue.
END_VAR
END_METHOD

{region 'Documentation'}
(*!
<summary>Restarts the script and resets the checking Assertions.</summary>
*)
{endregion}
METHOD PROTECTED ProcessReset
FStep := InitializeSubjects;
FChecked := FALSE;
FObservationReady := FALSE;
FExpectedObservationCount := 0;
FExpectedExplicitCount := 0;
FInitialization.Reset();
FInitializationMatches := TRUE;
FEnabled.Reset();
FEnabledMatches := TRUE;
FObservation.Reset();
FObservationMatches := TRUE;
FDirectEvaluation.Reset();
FDirectEvaluationMatches := TRUE;
FExplicitEvaluation.Reset();
FExplicitEvaluationMatches := TRUE;
FHookDispatch.Reset();
FHookDispatchMatches := TRUE;
FStableProperties.Reset();
FStablePropertiesMatches := TRUE;
FNoFindings.Reset();
FNoFindingsMatches := TRUE;
CompleteReset();
END_METHOD

{region 'Documentation'}
(*!
<summary>Advances one bounded script step per active PLC cycle.</summary>
*)
{endregion}
METHOD PROTECTED ProcessTests
VAR_INPUT
    Enable : BOOL; //! Phase permission supplied by the owning Test Case; FALSE does not authorize progression, while observation may continue.
END_VAR
IF NOT Enable THEN
    RETURN;
END_IF;
IF FChecked THEN
    FChecked := FALSE;
    FObservationReady := FALSE;
    IF FStep = ContinuedCall THEN
        CompleteTests();
        RETURN;
    END_IF;
    FStep := FStep + 1;
END_IF;
IF FStep = InitializeSubjects THEN
    InitializeActivitySubjects();
    RETURN;
END_IF;
SelectCall();
ObserveCall();
END_METHOD

{region 'Documentation'}
(*!
<summary>Selects literal inputs and expected gates for the current trace step.</summary>
*)
{endregion}
METHOD PRIVATE SelectCall
FEnable := FALSE;
FEvaluate := FALSE;
FExpectedObservation := FALSE;
FExpectedExplicitEvaluation := FALSE;
CASE FStep OF
    ConsumeInitialReset:
        FEnable := TRUE;
        FEvaluate := TRUE;
    DisabledCall:
        FEnable := FALSE;
    FirstEnabledCall, FirstReenabledCall:
        FEnable := TRUE;
        FEvaluate := TRUE;
        FExpectedObservation := ObserveFirstCycle;
        FExpectedExplicitEvaluation := TRUE;
    ObservationOnly:
        FEnable := TRUE;
        FExpectedObservation := TRUE;
    EvaluationOnly:
        FEvaluate := TRUE;
        FExpectedExplicitEvaluation := TRUE;
    ContinuedCall:
        FEnable := TRUE;
        FEvaluate := TRUE;
        FExpectedObservation := TRUE;
        FExpectedExplicitEvaluation := TRUE;
ELSE
    Error(Message := 'Unknown Assertion activity step.');
END_CASE;
END_METHOD

END_FUNCTION_BLOCK

// ---- SelfTests/TestCases/TestSuite_AssertionLifecycle/Helper/AssertionEvaluationSubject.TcPOU
{region 'Documentation'}
(*!
<summary>Exposes calls and activity gates of AssertionWithEvaluationBase without replacing its processing.</summary>
<description>
Bind the local publisher before Initialize. The inherited body owns initialization,
reset priority and activity history. Assert records both gates and a bounded sample;
active evaluation dispatches the selected inherited finding method without a result guard.
This deliberately exercises base-owned suppression. Counters are cumulative until ClearTrace.
ResetAssertion clears the sample and records the input available on the reset call.
The outer test owns expectations; this subject does not compute expected gates.
</description>
*)
{endregion}
FUNCTION_BLOCK AssertionEvaluationSubject EXTENDS AssertionWithEvaluationBase
VAR_INPUT
    Sample : UINT := 0; //! Controlled sample captured only while observation is active.
    Finding : E_Result := E_Result.Passed; //! Passed, Failed or Error finding dispatched only while evaluation is active.
    FindingMessage : STRING(GVL_Constants.MessageLength) := 'Controlled finding.'; //! Diagnostic text supplied to the selected Fail or Error operation.
END_VAR
VAR_OUTPUT
    AssertCallCount : UINT; //! Cumulative Assert-hook invocations since ClearTrace.
    ResetCallCount : UINT; //! Cumulative ResetAssertion-hook invocations since ClearTrace.
    ObservationCount : UINT; //! Cumulative Assert calls with the observation gate active since ClearTrace.
    EvaluationCount : UINT; //! Cumulative Assert calls with the evaluation gate active since ClearTrace.
    ObservedSample : UINT; //! Last Sample accepted while observation was active; ResetAssertion clears it.
    ResetSample : UINT; //! Sample present at the latest ResetAssertion call.
    ObservationDuringAssert : BOOL; //! Observation gate recorded on the latest Assert-hook entry.
    EvaluationDuringAssert : BOOL; //! Evaluation gate recorded on the latest Assert-hook entry.
END_VAR

SUPER^();

{region 'Documentation'}
(*!
<summary>Records inherited gates and evaluates only when permitted.</summary>
*)
{endregion}
METHOD PROTECTED Assert
AssertCallCount := AssertCallCount + 1;
ObservationDuringAssert := ObservationActive;
EvaluationDuringAssert := EvaluationActive;
IF ObservationDuringAssert THEN
    ObservationCount := ObservationCount + 1;
    ObservedSample := Sample;
END_IF;
IF EvaluationDuringAssert THEN
    EvaluationCount := EvaluationCount + 1;
    CASE Finding OF
        E_Result.Passed:
            Pass();
        E_Result.Failed:
            Fail(Message := FindingMessage);
        E_Result.Error:
            Error(Message := FindingMessage);
    ELSE
        RETURN;
    END_CASE;
END_IF;
END_METHOD

{region 'Documentation'}
(*!
<summary>Clears only test instrumentation; never changes inherited Assertion state.</summary>
*)
{endregion}
METHOD PUBLIC ClearTrace
AssertCallCount := 0;
ResetCallCount := 0;
ObservationCount := 0;
EvaluationCount := 0;
ObservedSample := 0;
ResetSample := 0;
ObservationDuringAssert := FALSE;
EvaluationDuringAssert := FALSE;
END_METHOD

{region 'Documentation'}
(*!
<summary>Records one reset with bound inputs and clears the observation sample.</summary>
*)
{endregion}
METHOD PROTECTED ResetAssertion
ResetCallCount := ResetCallCount + 1;
ResetSample := Sample;
ObservedSample := 0;
END_METHOD

END_FUNCTION_BLOCK

// ---- Framework/Assertions/POU/AssertionWithEvaluationBase.TcPOU
{region 'Documentation'}
(*!
<summary>Base for observation and explicitly requested result evaluation.</summary>
<description>

Enable and ObserveFirstCycle control ObservationActive. Evaluate controls
EvaluationActive independently of both, provided initialization succeeded and this is not a
reset call. Evaluate is a level input, not a latched request.

A concrete Assert implementation performs observation under ObservationActive and decides
the held result under EvaluationActive. Evaluation with Enable FALSE is supported;
ObserveFirstCycle delays observation, not explicit evaluation. Derived FB bodies call SUPER^()
once.

</description>
*)
{endregion}
FUNCTION_BLOCK ABSTRACT AssertionWithEvaluationBase EXTENDS AssertionBase
VAR_INPUT
    Evaluate : BOOL; //! Requests result evaluation independently of Enable; initialization and reset still gate evaluation.
END_VAR
VAR
    FEvaluate : BOOL;
END_VAR

FEvaluate := Evaluate;
SUPER^();

{region 'Documentation'}
(*!
<summary>Indicate explicit evaluation independently of observation.</summary>
<description>

TRUE when initialized, Evaluate was accepted by the FB call and the call is not
resetting. Neither Enable nor ObserveFirstCycle suppresses this gate.

</description>
*)
{endregion}
{attribute 'monitoring' := 'call'}
PROPERTY PUBLIC EvaluationActive : BOOL //! TRUE when initialized, Evaluate was accepted and the call is not resetting; independent of Enable.
GET // PUBLIC
EvaluationActive := IsInitialized AND FEvaluate AND NOT FResetActive;
END_GET
END_PROPERTY

END_FUNCTION_BLOCK

// ---- SelfTests/TestCases/TestSuite_AssertionLifecycle/Test_AssertionUninitialized.TcPOU
{region 'Documentation'}
(*!
<summary>Checks that both Assertion bases remain passive before Initialize.</summary>
<description>
Neither subject is initialized. Calls request observation and evaluation deliberately.
The same uninitialized instances are reused after outer Reset, without rewriting
production state. Instrumentation is cleared separately from the inherited state.
</description>
*)
{endregion}
FUNCTION_BLOCK Test_AssertionUninitialized EXTENDS TestCaseBase
VAR
    FDirect : AssertionLifecycleSubject;
    FExplicit : AssertionEvaluationSubject;
    FCapture : EventBuffer;
    FEvents : ARRAY[1..CaptureLength] OF ST_Event;
    FCaptureFifo : ST_FifoStatus;
    FCaptureStatus : ST_EventBufferStatus;
    FCallCount : UINT;
    FObservationReady : BOOL;
    FChecked : BOOL;
END_VAR
VAR
    FPassiveState : AssertTrue;
    FPassiveStateMatches : BOOL;
    FNoHooks : AssertTrue;
    FNoHooksMatches : BOOL;
    FNoFindings : AssertTrue;
    FNoFindingsMatches : BOOL;
END_VAR
VAR CONSTANT
    CaptureLength : UINT := 8;
    ObservationCalls : UINT := 2;
END_VAR

SUPER^();

{region 'Documentation'}
(*!
<summary>Collects only outer checking Assertions, never intentional subject findings.</summary>
*)
{endregion}
METHOD PROTECTED AggregateResults
VAR_INPUT
    Aggregator : I_ResultAggregator; //! Borrowed result sink owned by the outer Test Case; add this test's checking Assertions without resetting or retaining the sink.
END_VAR
Aggregator.AddProvider(Provider := FPassiveState);
Aggregator.AddProvider(Provider := FNoHooks);
Aggregator.AddProvider(Provider := FNoFindings);
END_METHOD

{region 'Documentation'}
(*!
<summary>Configures checking Assertions; subject actions remain in the test script.</summary>
*)
{endregion}
METHOD PROTECTED Configure
FPreparationStateCount := 0;
FTestStateCount := 1;
FPassiveState.Initialize(Parent := THIS^,
    AssertionName := 'PassiveState');
FNoHooks.Initialize(Parent := THIS^,
    AssertionName := 'NoHooks');
FNoFindings.Initialize(Parent := THIS^,
    AssertionName := 'NoFindings');
FDirect.BindPublisher(Publisher := FCapture);
FExplicit.BindPublisher(Publisher := FCapture);
END_METHOD

{region 'Documentation'}
(*!
<summary>Completes abort without asynchronous resources.</summary>
*)
{endregion}
METHOD PROTECTED ProcessAbort
VAR_INPUT
    Enable : BOOL; //! Phase permission supplied by the owning Test Case; FALSE does not authorize progression, while observation may continue.
END_VAR
IF Enable THEN
    CompleteAbort();
END_IF;
END_METHOD

{region 'Documentation'}
(*!
<summary>Latches checked observations before the next script step may proceed.</summary>
*)
{endregion}
METHOD PROTECTED ProcessAssertions
VAR_INPUT
    Enable : BOOL; //! Phase permission supplied by the owning Test Case; FALSE does not authorize progression, while observation may continue.
END_VAR
VAR
    Evaluate : BOOL;
END_VAR
Evaluate := Enable AND FObservationReady;
FPassiveState(Enable := Evaluate,
    State := State,
    IN := FPassiveStateMatches);
FNoHooks(Enable := Evaluate,
    State := State,
    IN := FNoHooksMatches);
FNoFindings(Enable := Evaluate,
    State := State,
    IN := FNoFindingsMatches);
IF Evaluate THEN
    FChecked := TRUE;
END_IF;
END_METHOD

{region 'Documentation'}
(*!
<summary>No Preparation phase is required.</summary>
*)
{endregion}
METHOD PROTECTED ProcessPreparations
VAR_INPUT
    // SA0033: Required hook; this test has no Preparation phase.
    {attribute 'analysis' := '-33'}
    Enable : BOOL; //! Phase permission supplied by the owning Test Case; FALSE does not authorize progression, while observation may continue.
END_VAR
END_METHOD

{region 'Documentation'}
(*!
<summary>Restarts the script and resets the checking Assertions.</summary>
*)
{endregion}
METHOD PROTECTED ProcessReset
FCallCount := 0;
FChecked := FALSE;
FObservationReady := FALSE;
FDirect.ClearTrace();
FExplicit.ClearTrace();
FPassiveState.Reset();
FPassiveStateMatches := TRUE;
FNoHooks.Reset();
FNoHooksMatches := TRUE;
FNoFindings.Reset();
FNoFindingsMatches := TRUE;
CompleteReset();
END_METHOD

{region 'Documentation'}
(*!
<summary>Advances one bounded script step per active PLC cycle.</summary>
*)
{endregion}
METHOD PROTECTED ProcessTests
VAR_INPUT
    Enable : BOOL; //! Phase permission supplied by the owning Test Case; FALSE does not authorize progression, while observation may continue.
END_VAR
IF NOT Enable THEN
    RETURN;
END_IF;
IF FChecked THEN
    FChecked := FALSE;
    FObservationReady := FALSE;
    IF FCallCount = ObservationCalls THEN
        CompleteTests();
        RETURN;
    END_IF;
END_IF;
IF FCallCount = 0 THEN
    IF NOT FCapture.Initialize(Buffer := FEvents,
        FifoControl := FCaptureFifo,
        Status := FCaptureStatus) THEN
        Error(Message := 'Uninitialized Assertion capture setup failed.');
        RETURN;
    END_IF;
END_IF;
FDirect(Enable := TRUE,
    State := E_State.Running);
FExplicit(Enable := TRUE,
    Evaluate := TRUE,
    State := E_State.Running);
FCallCount := FCallCount + 1;
FPassiveStateMatches := NOT FDirect.IsInitialized AND NOT FExplicit.IsInitialized
    AND FDirect.Enabled AND FExplicit.Enabled
    AND NOT FDirect.ObservationActive AND NOT FExplicit.ObservationActive
    AND NOT FDirect.EvaluationActive AND NOT FExplicit.EvaluationActive
    AND (FDirect.Result = E_Result.NotEvaluated) AND (FExplicit.Result = E_Result.NotEvaluated);
FNoHooksMatches := (FDirect.AssertCallCount = 0) AND (FExplicit.AssertCallCount = 0)
    AND (FDirect.ResetCallCount = 0) AND (FExplicit.ResetCallCount = 0);
FNoFindingsMatches := (FCaptureStatus.SequenceId = 0) AND (FCaptureStatus.LostEventCount = 0);
FObservationReady := TRUE;
END_METHOD

END_FUNCTION_BLOCK

// ---- SelfTests/TestCases/TestSuite_AssertionLifecycle/Test_AssertionResetReuse.TcPOU
{region 'Documentation'}
(*!
<summary>Checks deferred reset priority and reuse for both Assertion bases.</summary>
<description>
The subject reset request is inspected before any subsequent FB call. Two requests
must coalesce into one reset hook. Reset retains identity/settings and suppresses
findings despite active inputs. Both subjects use ObserveFirstCycle FALSE, so the
first enabled call after reset must still be excluded. Each subject emits one Failed
finding before reset and one after reset; repeated failure must not emit another.
</description>
*)
{endregion}
FUNCTION_BLOCK Test_AssertionResetReuse EXTENDS TestCaseBase
VAR
    FDirect : AssertionLifecycleSubject;
    FExplicit : AssertionEvaluationSubject;
    FCapture : EventBuffer;
    FEvents : ARRAY[1..CaptureLength] OF ST_Event;
    FCaptureFifo : ST_FifoStatus;
    FCaptureStatus : ST_EventBufferStatus;
    FStep : UINT;
    FChecked : BOOL;
    FObservationReady : BOOL;
END_VAR
VAR
    FDeferredReset : AssertTrue;
    FDeferredResetMatches : BOOL;
    FResetPriority : AssertTrue;
    FResetPriorityMatches : BOOL;
    FHookDispatch : AssertTrue;
    FHookDispatchMatches : BOOL;
    FFirstObservation : AssertTrue;
    FFirstObservationMatches : BOOL;
    FRetainedResult : AssertTrue;
    FRetainedResultMatches : BOOL;
    FConfiguration : AssertTrue;
    FConfigurationMatches : BOOL;
    FFindings : AssertTrue;
    FFindingsMatches : BOOL;
    FCaptureIntegrity : AssertTrue;
    FCaptureIntegrityMatches : BOOL;
END_VAR
VAR CONSTANT
    CaptureLength : UINT := 16;
    InitializeSubjects : UINT := 0;
    InitialReset : UINT := 1;
    FirstEnable : UINT := 2;
    ProduceFailure : UINT := 3;
    DisabledHolding : UINT := 4;
    RequestTwice : UINT := 5;
    ConsumeReset : UINT := 6;
    FirstEnableAfterReset : UINT := 7;
    FailureAfterReset : UINT := 8;
    RepeatedFailure : UINT := 9;
    SampleBeforeReset : UINT := 23;
    SampleAtReset : UINT := 41;
    SampleAfterReset : UINT := 67;
END_VAR

SUPER^();

{region 'Documentation'}
(*!
<summary>Collects only outer checking Assertions, never intentional subject findings.</summary>
*)
{endregion}
METHOD PROTECTED AggregateResults
VAR_INPUT
    Aggregator : I_ResultAggregator; //! Borrowed result sink owned by the outer Test Case; add this test's checking Assertions without resetting or retaining the sink.
END_VAR
Aggregator.AddProvider(Provider := FDeferredReset);
Aggregator.AddProvider(Provider := FResetPriority);
Aggregator.AddProvider(Provider := FHookDispatch);
Aggregator.AddProvider(Provider := FFirstObservation);
Aggregator.AddProvider(Provider := FRetainedResult);
Aggregator.AddProvider(Provider := FConfiguration);
Aggregator.AddProvider(Provider := FFindings);
Aggregator.AddProvider(Provider := FCaptureIntegrity);
END_METHOD

{region 'Documentation'}
(*!
<summary>Calls each subject once with the same controlled failed finding.</summary>
*)
{endregion}
METHOD PRIVATE CallSubjects
VAR_INPUT
    Enable : BOOL; //! Observation-enable input forwarded to the controlled Assertion subjects for this call.
    Evaluate : BOOL; //! Explicit evaluation request forwarded to the evaluation-gated subjects.
    Sample : UINT; //! Controlled sample forwarded to all subjects for this call.
END_VAR
FDirect(Enable := Enable,
    State := E_State.Running,
    Sample := Sample,
    Finding := E_Result.Failed);
FExplicit(Enable := Enable,
    Evaluate := Evaluate,
    State := E_State.Running,
    Sample := Sample,
    Finding := E_Result.Failed);
END_METHOD

{region 'Documentation'}
(*!
<summary>Checks that ordinary Reset preserves identity, initialization and settings.</summary>
*)
{endregion}
METHOD PRIVATE CheckConfiguration
FConfigurationMatches := FDirect.IsInitialized AND FExplicit.IsInitialized
    AND (FDirect.Name = CONCAT(Name, '.DirectSubject'))
    AND (FExplicit.Name = CONCAT(Name, '.ExplicitSubject'))
    AND (FDirect.ResourceName = 'DirectResource')
    AND (FExplicit.ResourceName = 'ExplicitResource')
    AND NOT FDirect.ObserveFirstCycle AND NOT FExplicit.ObserveFirstCycle;
END_METHOD

{region 'Documentation'}
(*!
<summary>Configures checking Assertions; subject actions remain in the test script.</summary>
*)
{endregion}
METHOD PROTECTED Configure
FPreparationStateCount := 0;
FTestStateCount := 1;
FDeferredReset.Initialize(Parent := THIS^,
    AssertionName := 'DeferredReset');
FResetPriority.Initialize(Parent := THIS^,
    AssertionName := 'ResetPriority');
FHookDispatch.Initialize(Parent := THIS^,
    AssertionName := 'HookDispatch');
FFirstObservation.Initialize(Parent := THIS^,
    AssertionName := 'FirstObservation');
FRetainedResult.Initialize(Parent := THIS^,
    AssertionName := 'RetainedResult');
FConfiguration.Initialize(Parent := THIS^,
    AssertionName := 'Configuration');
FFindings.Initialize(Parent := THIS^,
    AssertionName := 'Findings');
FCaptureIntegrity.Initialize(Parent := THIS^,
    AssertionName := 'CaptureIntegrity');
FDirect.BindPublisher(Publisher := FCapture);
FExplicit.BindPublisher(Publisher := FCapture);
END_METHOD

{region 'Documentation'}
(*!
<summary>Establishes fresh configured subjects for each outer test run.</summary>
*)
{endregion}
METHOD PRIVATE InitializeResetSubjects
VAR
    DirectInitialized : BOOL;
    ExplicitInitialized : BOOL;
END_VAR
IF NOT FCapture.Initialize(Buffer := FEvents,
    FifoControl := FCaptureFifo,
    Status := FCaptureStatus) THEN
    Error(Message := 'Assertion reset capture setup failed.');
    RETURN;
END_IF;
FDirect.ClearTrace();
FExplicit.ClearTrace();
DirectInitialized := FDirect.Initialize(Parent := THIS^,
    AssertionName := 'DirectSubject',
    ResourceName := 'DirectResource',
    ObserveFirstCycle := FALSE);
ExplicitInitialized := FExplicit.Initialize(Parent := THIS^,
    AssertionName := 'ExplicitSubject',
    ResourceName := 'ExplicitResource',
    ObserveFirstCycle := FALSE);
IF NOT DirectInitialized OR NOT ExplicitInitialized THEN
    Error(Message := 'Assertion reset subjects could not be initialized.');
    RETURN;
END_IF;
FStep := InitialReset;
END_METHOD

{region 'Documentation'}
(*!
<summary>Completes abort without asynchronous resources.</summary>
*)
{endregion}
METHOD PROTECTED ProcessAbort
VAR_INPUT
    Enable : BOOL; //! Phase permission supplied by the owning Test Case; FALSE does not authorize progression, while observation may continue.
END_VAR
IF Enable THEN
    CompleteAbort();
END_IF;
END_METHOD

{region 'Documentation'}
(*!
<summary>Latches checked observations before the next script step may proceed.</summary>
*)
{endregion}
METHOD PROTECTED ProcessAssertions
VAR_INPUT
    Enable : BOOL; //! Phase permission supplied by the owning Test Case; FALSE does not authorize progression, while observation may continue.
END_VAR
VAR
    Evaluate : BOOL;
END_VAR
Evaluate := Enable AND FObservationReady;
FDeferredReset(Enable := Evaluate,
    State := State,
    IN := FDeferredResetMatches);
FResetPriority(Enable := Evaluate,
    State := State,
    IN := FResetPriorityMatches);
FHookDispatch(Enable := Evaluate,
    State := State,
    IN := FHookDispatchMatches);
FFirstObservation(Enable := Evaluate,
    State := State,
    IN := FFirstObservationMatches);
FRetainedResult(Enable := Evaluate,
    State := State,
    IN := FRetainedResultMatches);
FConfiguration(Enable := Evaluate,
    State := State,
    IN := FConfigurationMatches);
FFindings(Enable := Evaluate,
    State := State,
    IN := FFindingsMatches);
FCaptureIntegrity(Enable := Evaluate,
    State := State,
    IN := FCaptureIntegrityMatches);
IF Evaluate THEN
    FChecked := TRUE;
END_IF;
END_METHOD

{region 'Documentation'}
(*!
<summary>No Preparation phase is required.</summary>
*)
{endregion}
METHOD PROTECTED ProcessPreparations
VAR_INPUT
    // SA0033: Required hook; this test has no Preparation phase.
    {attribute 'analysis' := '-33'}
    Enable : BOOL; //! Phase permission supplied by the owning Test Case; FALSE does not authorize progression, while observation may continue.
END_VAR
END_METHOD

{region 'Documentation'}
(*!
<summary>Restarts the script and resets the checking Assertions.</summary>
*)
{endregion}
METHOD PROTECTED ProcessReset
FStep := InitializeSubjects;
FChecked := FALSE;
FObservationReady := FALSE;
FDeferredReset.Reset();
FDeferredResetMatches := TRUE;
FResetPriority.Reset();
FResetPriorityMatches := TRUE;
FHookDispatch.Reset();
FHookDispatchMatches := TRUE;
FFirstObservation.Reset();
FFirstObservationMatches := TRUE;
FRetainedResult.Reset();
FRetainedResultMatches := TRUE;
FConfiguration.Reset();
FConfigurationMatches := TRUE;
FFindings.Reset();
FFindingsMatches := TRUE;
FCaptureIntegrity.Reset();
FCaptureIntegrityMatches := TRUE;
CompleteReset();
END_METHOD

{region 'Documentation'}
(*!
<summary>Advances one bounded script step per active PLC cycle.</summary>
*)
{endregion}
METHOD PROTECTED ProcessTests
VAR_INPUT
    Enable : BOOL; //! Phase permission supplied by the owning Test Case; FALSE does not authorize progression, while observation may continue.
END_VAR
IF NOT Enable THEN
    RETURN;
END_IF;
IF FChecked THEN
    FChecked := FALSE;
    FObservationReady := FALSE;
    IF FStep = RepeatedFailure THEN
        CompleteTests();
        RETURN;
    END_IF;
    FStep := FStep + 1;
END_IF;
IF FStep = InitializeSubjects THEN
    InitializeResetSubjects();
    RETURN;
END_IF;
RunStep();
CheckConfiguration();
FObservationReady := TRUE;
END_METHOD

{region 'Documentation'}
(*!
<summary>Runs one reset/reuse operation and records independent expected observations.</summary>
*)
{endregion}
METHOD PRIVATE RunStep
CASE FStep OF
    InitialReset:
        CallSubjects(Enable := TRUE,
            Evaluate := TRUE,
            Sample := SampleAtReset);
        FResetPriorityMatches := (FDirect.Result = E_Result.NotEvaluated)
            AND (FExplicit.Result = E_Result.NotEvaluated)
            AND NOT FDirect.ObservationActive AND NOT FExplicit.ObservationActive
            AND NOT FDirect.EvaluationActive AND NOT FExplicit.EvaluationActive;
        FHookDispatchMatches := (FDirect.ResetCallCount = 1) AND (FExplicit.ResetCallCount = 1)
            AND (FDirect.AssertCallCount = 0) AND (FExplicit.AssertCallCount = 0);
        FFindingsMatches := FCaptureStatus.SequenceId = 0;
    FirstEnable, FirstEnableAfterReset:
        CallSubjects(Enable := TRUE,
            Evaluate := FALSE,
            Sample := SampleBeforeReset);
        FFirstObservationMatches := NOT FDirect.ObservationActive AND NOT FExplicit.ObservationActive
            AND NOT FDirect.EvaluationActive AND NOT FExplicit.EvaluationActive
            AND (FDirect.ObservedSample = 0) AND (FExplicit.ObservedSample = 0)
            AND (FDirect.Result = E_Result.NotEvaluated) AND (FExplicit.Result = E_Result.NotEvaluated);
    ProduceFailure:
        CallSubjects(Enable := TRUE,
            Evaluate := TRUE,
            Sample := SampleBeforeReset);
        FRetainedResultMatches := (FDirect.Result = E_Result.Failed)
            AND (FExplicit.Result = E_Result.Failed);
        FFindingsMatches := FCaptureStatus.SequenceId = 2;
    DisabledHolding:
        CallSubjects(Enable := FALSE,
            Evaluate := FALSE,
            Sample := SampleAtReset);
        FRetainedResultMatches := (FDirect.Result = E_Result.Failed)
            AND (FExplicit.Result = E_Result.Failed)
            AND (FDirect.ObservedSample = SampleBeforeReset)
            AND (FExplicit.ObservedSample = SampleBeforeReset);
        FFindingsMatches := FCaptureStatus.SequenceId = 2;
    RequestTwice:
        FDirect.Reset();
        FDirect.Reset();
        FExplicit.Reset();
        FExplicit.Reset();
        FDeferredResetMatches := (FDirect.Result = E_Result.Failed)
            AND (FExplicit.Result = E_Result.Failed)
            AND (FDirect.ObservedSample = SampleBeforeReset)
            AND (FExplicit.ObservedSample = SampleBeforeReset)
            AND (FDirect.ResetCallCount = 1) AND (FExplicit.ResetCallCount = 1);
        FFindingsMatches := FCaptureStatus.SequenceId = 2;
    ConsumeReset:
        CallSubjects(Enable := TRUE,
            Evaluate := TRUE,
            Sample := SampleAtReset);
        FResetPriorityMatches := (FDirect.Result = E_Result.NotEvaluated)
            AND (FExplicit.Result = E_Result.NotEvaluated)
            AND NOT FDirect.ObservationActive AND NOT FExplicit.ObservationActive
            AND NOT FDirect.EvaluationActive AND NOT FExplicit.EvaluationActive;
        FHookDispatchMatches := (FDirect.ResetCallCount = 2) AND (FExplicit.ResetCallCount = 2)
            AND (FDirect.AssertCallCount = 3) AND (FExplicit.AssertCallCount = 3)
            AND (FDirect.ResetSample = SampleAtReset) AND (FExplicit.ResetSample = SampleAtReset)
            AND (FDirect.ObservedSample = 0) AND (FExplicit.ObservedSample = 0);
        FFindingsMatches := FCaptureStatus.SequenceId = 2;
    FailureAfterReset, RepeatedFailure:
        CallSubjects(Enable := TRUE,
            Evaluate := TRUE,
            Sample := SampleAfterReset);
        FRetainedResultMatches := (FDirect.Result = E_Result.Failed)
            AND (FExplicit.Result = E_Result.Failed)
            AND (FDirect.ObservedSample = SampleAfterReset)
            AND (FExplicit.ObservedSample = SampleAfterReset);
        FFindingsMatches := FCaptureStatus.SequenceId = 4;
ELSE
    Error(Message := 'Unknown Assertion reset step.');
END_CASE;
FCaptureIntegrityMatches := FCaptureStatus.LostEventCount = 0;
END_METHOD

END_FUNCTION_BLOCK

// ---- SelfTests/TestCases/TestSuite_AssertionLifecycle/Test_AssertionEscalation.TcPOU
{region 'Documentation'}
(*!
<summary>Checks monotonic Assertion results and transition-only event publication.</summary>
<description>
A controlled concrete Assert dispatches each selected protected finding method even
when the result is already Failed or Error. No subject guard can mask a broken base
suppression rule. The first epoch checks all attempted downgrades; two reset epochs
check direct NotEvaluated-to-Failed and NotEvaluated-to-Error. Each step checks the
held result and exact event count. The final check inspects all four finding payloads.
</description>
*)
{endregion}
FUNCTION_BLOCK Test_AssertionEscalation EXTENDS TestCaseBase
VAR
    FSubject : AssertionLifecycleSubject;
    FCapture : EventBuffer;
    FEvents : ARRAY[1..CaptureLength] OF ST_Event;
    FCaptureFifo : ST_FifoStatus;
    FCaptureStatus : ST_EventBufferStatus;
    FStep : UINT;
    FChecked : BOOL;
    FObservationReady : BOOL;
    FFinding : E_Result;
    FExpectedResult : E_Result;
    FExpectedEvents : UDINT;
    FMessage : STRING(GVL_Constants.MessageLength);
END_VAR
VAR
    FResultPriority : AssertTrue;
    FResultPriorityMatches : BOOL;
    FFindingCount : AssertTrue;
    FFindingCountMatches : BOOL;
    FFindingPayload : AssertTrue;
    FFindingPayloadMatches : BOOL;
    FCaptureIntegrity : AssertTrue;
    FCaptureIntegrityMatches : BOOL;
END_VAR
VAR CONSTANT
    CaptureLength : UINT := 16;
    InitializeSubject : UINT := 0;
    InitialReset : UINT := 1;
    PassInitially : UINT := 2;
    RepeatPass : UINT := 3;
    FailAfterPass : UINT := 4;
    RepeatFail : UINT := 5;
    PassAfterFail : UINT := 6;
    ErrorAfterFail : UINT := 7;
    RepeatError : UINT := 8;
    FailAfterError : UINT := 9;
    PassAfterError : UINT := 10;
    ResetForDirectFail : UINT := 11;
    DirectFail : UINT := 12;
    ResetForDirectError : UINT := 13;
    DirectError : UINT := 14;
    RepeatDirectError : UINT := 15;
END_VAR

SUPER^();

{region 'Documentation'}
(*!
<summary>Collects only outer checking Assertions, never intentional subject findings.</summary>
*)
{endregion}
METHOD PROTECTED AggregateResults
VAR_INPUT
    Aggregator : I_ResultAggregator; //! Borrowed result sink owned by the outer Test Case; add this test's checking Assertions without resetting or retaining the sink.
END_VAR
Aggregator.AddProvider(Provider := FResultPriority);
Aggregator.AddProvider(Provider := FFindingCount);
Aggregator.AddProvider(Provider := FFindingPayload);
Aggregator.AddProvider(Provider := FCaptureIntegrity);
END_METHOD

{region 'Documentation'}
(*!
<summary>Checks the four retained findings against fixed expected context and classifications.</summary>
*)
{endregion}
METHOD PRIVATE CheckFindingPayloads
VAR
    Index : UINT;
    ExpectedResult : E_Result;
    ExpectedSeverity : E_EventSeverity;
    ExpectedMessage : STRING(GVL_Constants.MessageLength);
END_VAR
FFindingPayloadMatches := TRUE;
FOR Index := 1 TO 4 DO
    CASE Index OF
        1, 3:
            ExpectedResult := E_Result.Failed;
            ExpectedSeverity := E_EventSeverity.Info;
            ExpectedMessage := 'Controlled Failed.';
        2, 4:
            ExpectedResult := E_Result.Error;
            ExpectedSeverity := E_EventSeverity.Error;
            ExpectedMessage := 'Controlled Error.';
    ELSE
        FFindingPayloadMatches := FALSE;
        RETURN;
    END_CASE;
    FFindingPayloadMatches := FFindingPayloadMatches
        AND (FEvents[Index].SequenceId = Index)
        AND (FEvents[Index].OwnerScope = E_OwnerScope.Assertion)
        AND (FEvents[Index].EventType = E_EventType.Result)
        AND (FEvents[Index].Severity = ExpectedSeverity)
        AND (FEvents[Index].Name = CONCAT(Name, '.Subject'))
        AND (FEvents[Index].ResourceName = 'ObservedResource')
        AND (FEvents[Index].State = E_State.Running)
        AND (FEvents[Index].Result = ExpectedResult)
        AND (FEvents[Index].Message = ExpectedMessage);
END_FOR;
END_METHOD

{region 'Documentation'}
(*!
<summary>Configures checking Assertions; subject actions remain in the test script.</summary>
*)
{endregion}
METHOD PROTECTED Configure
FPreparationStateCount := 0;
FTestStateCount := 1;
FResultPriority.Initialize(Parent := THIS^,
    AssertionName := 'ResultPriority');
FFindingCount.Initialize(Parent := THIS^,
    AssertionName := 'FindingCount');
FFindingPayload.Initialize(Parent := THIS^,
    AssertionName := 'FindingPayload');
FCaptureIntegrity.Initialize(Parent := THIS^,
    AssertionName := 'CaptureIntegrity');
FSubject.BindPublisher(Publisher := FCapture);
END_METHOD

{region 'Documentation'}
(*!
<summary>Starts a fresh subject run without clearing evidence between its reset epochs.</summary>
*)
{endregion}
METHOD PRIVATE InitializeEscalationSubject
IF NOT FCapture.Initialize(Buffer := FEvents,
    FifoControl := FCaptureFifo,
    Status := FCaptureStatus) THEN
    Error(Message := 'Assertion escalation capture setup failed.');
    RETURN;
END_IF;
IF NOT FSubject.Initialize(Parent := THIS^,
    AssertionName := 'Subject',
    ResourceName := 'ObservedResource') THEN
    Error(Message := 'Assertion escalation subject initialization failed.');
    RETURN;
END_IF;
FStep := InitialReset;
END_METHOD

{region 'Documentation'}
(*!
<summary>Completes abort without asynchronous resources.</summary>
*)
{endregion}
METHOD PROTECTED ProcessAbort
VAR_INPUT
    Enable : BOOL; //! Phase permission supplied by the owning Test Case; FALSE does not authorize progression, while observation may continue.
END_VAR
IF Enable THEN
    CompleteAbort();
END_IF;
END_METHOD

{region 'Documentation'}
(*!
<summary>Latches checked observations before the next script step may proceed.</summary>
*)
{endregion}
METHOD PROTECTED ProcessAssertions
VAR_INPUT
    Enable : BOOL; //! Phase permission supplied by the owning Test Case; FALSE does not authorize progression, while observation may continue.
END_VAR
VAR
    Evaluate : BOOL;
END_VAR
Evaluate := Enable AND FObservationReady;
FResultPriority(Enable := Evaluate,
    State := State,
    IN := FResultPriorityMatches);
FFindingCount(Enable := Evaluate,
    State := State,
    IN := FFindingCountMatches);
FFindingPayload(Enable := Evaluate,
    State := State,
    IN := FFindingPayloadMatches);
FCaptureIntegrity(Enable := Evaluate,
    State := State,
    IN := FCaptureIntegrityMatches);
IF Evaluate THEN
    FChecked := TRUE;
END_IF;
END_METHOD

{region 'Documentation'}
(*!
<summary>No Preparation phase is required.</summary>
*)
{endregion}
METHOD PROTECTED ProcessPreparations
VAR_INPUT
    // SA0033: Required hook; this test has no Preparation phase.
    {attribute 'analysis' := '-33'}
    Enable : BOOL; //! Phase permission supplied by the owning Test Case; FALSE does not authorize progression, while observation may continue.
END_VAR
END_METHOD

{region 'Documentation'}
(*!
<summary>Restarts the script and resets the checking Assertions.</summary>
*)
{endregion}
METHOD PROTECTED ProcessReset
FStep := InitializeSubject;
FChecked := FALSE;
FObservationReady := FALSE;
FResultPriority.Reset();
FResultPriorityMatches := TRUE;
FFindingCount.Reset();
FFindingCountMatches := TRUE;
FFindingPayload.Reset();
FFindingPayloadMatches := TRUE;
FCaptureIntegrity.Reset();
FCaptureIntegrityMatches := TRUE;
CompleteReset();
END_METHOD

{region 'Documentation'}
(*!
<summary>Advances one bounded script step per active PLC cycle.</summary>
*)
{endregion}
METHOD PROTECTED ProcessTests
VAR_INPUT
    Enable : BOOL; //! Phase permission supplied by the owning Test Case; FALSE does not authorize progression, while observation may continue.
END_VAR
IF NOT Enable THEN
    RETURN;
END_IF;
IF FChecked THEN
    FChecked := FALSE;
    FObservationReady := FALSE;
    IF FStep = RepeatDirectError THEN
        CompleteTests();
        RETURN;
    END_IF;
    FStep := FStep + 1;
END_IF;
IF FStep = InitializeSubject THEN
    InitializeEscalationSubject();
    RETURN;
END_IF;
SelectFinding();
IF FFinding = E_Result.Error THEN
    FMessage := 'Controlled Error.';
ELSE
    FMessage := 'Controlled Failed.';
END_IF;
FSubject(Enable := TRUE,
    State := E_State.Running,
    Finding := FFinding,
    FindingMessage := FMessage);
FResultPriorityMatches := FSubject.Result = FExpectedResult;
FFindingCountMatches := FCaptureStatus.SequenceId = FExpectedEvents;
FCaptureIntegrityMatches := FCaptureStatus.LostEventCount = 0;
IF FStep = RepeatDirectError THEN
    CheckFindingPayloads();
END_IF;
FObservationReady := TRUE;
END_METHOD

{region 'Documentation'}
(*!
<summary>Selects explicit finding attempts, held-result expectations and exact event totals.</summary>
*)
{endregion}
METHOD PRIVATE SelectFinding
CASE FStep OF
    InitialReset:
        FFinding := E_Result.Error;
        FExpectedResult := E_Result.NotEvaluated;
        FExpectedEvents := 0;
    PassInitially:
        FFinding := E_Result.Passed;
        FExpectedResult := E_Result.Passed;
        FExpectedEvents := 0;
    RepeatPass:
        FFinding := E_Result.Passed;
        FExpectedResult := E_Result.Passed;
        FExpectedEvents := 0;
    FailAfterPass:
        FFinding := E_Result.Failed;
        FExpectedResult := E_Result.Failed;
        FExpectedEvents := 1;
    RepeatFail:
        FFinding := E_Result.Failed;
        FExpectedResult := E_Result.Failed;
        FExpectedEvents := 1;
    PassAfterFail:
        FFinding := E_Result.Passed;
        FExpectedResult := E_Result.Failed;
        FExpectedEvents := 1;
    ErrorAfterFail:
        FFinding := E_Result.Error;
        FExpectedResult := E_Result.Error;
        FExpectedEvents := 2;
    RepeatError:
        FFinding := E_Result.Error;
        FExpectedResult := E_Result.Error;
        FExpectedEvents := 2;
    FailAfterError:
        FFinding := E_Result.Failed;
        FExpectedResult := E_Result.Error;
        FExpectedEvents := 2;
    PassAfterError:
        FFinding := E_Result.Passed;
        FExpectedResult := E_Result.Error;
        FExpectedEvents := 2;
    ResetForDirectFail:
        FSubject.Reset();
        FFinding := E_Result.Error;
        FExpectedResult := E_Result.NotEvaluated;
        FExpectedEvents := 2;
    DirectFail:
        FFinding := E_Result.Failed;
        FExpectedResult := E_Result.Failed;
        FExpectedEvents := 3;
    ResetForDirectError:
        FSubject.Reset();
        FFinding := E_Result.Error;
        FExpectedResult := E_Result.NotEvaluated;
        FExpectedEvents := 3;
    DirectError:
        FFinding := E_Result.Error;
        FExpectedResult := E_Result.Error;
        FExpectedEvents := 4;
    RepeatDirectError:
        FFinding := E_Result.Error;
        FExpectedResult := E_Result.Error;
        FExpectedEvents := 4;
ELSE
    Error(Message := 'Unknown Assertion escalation step.');
END_CASE;
END_METHOD

END_FUNCTION_BLOCK

// ---- SelfTests/TestSuites/TestSuite_AssertionComparisons.TcPOU
{region 'Documentation'}
(*!
<summary>Checks scalar comparisons, ranges, temporal boundaries and diagnostic rendering.</summary>
*)
{endregion}
FUNCTION_BLOCK TestSuite_AssertionComparisons EXTENDS TestSuiteBase
VAR
    FSignedRelations : Test_AssertionSignedRelations;
    FUnsignedRelations : Test_AssertionUnsignedRelations;
    FBitEquality : Test_AssertionBitEquality;
    FBooleanComparisons : Test_AssertionBooleanComparisons;
    FCharacterEquality : Test_AssertionCharacterEquality;
    FSignedRanges : Test_AssertionSignedRanges;
    FUnsignedRanges : Test_AssertionUnsignedRanges;
    FDurationComparisons : Test_AssertionDurationComparisons;
    FDateNormalization : Test_AssertionDateNormalization;
    FTODDomain : Test_AssertionTODDomain;
    FLTODDomain : Test_AssertionLTODDomain;
    FScalarDiagnostics : Test_AssertionScalarDiagnostics;
    FTestCases : ARRAY[1..TestCaseCapacity] OF I_TestCase;
END_VAR
VAR CONSTANT
    TestCaseCapacity : UINT := 12;
END_VAR

SUPER^();

{region 'Documentation'}
(*!
<summary>Initializes and registers the twelve isolated scalar comparison scenarios.</summary>
*)
{endregion}
METHOD PROTECTED Configure
VAR_IN_OUT
    // SA0167: Borrowed owner builder; no temporary instance is created.
    {attribute 'analysis' := '-167'}
    Builder : TestSuiteConfigurationBuilder; //! Borrowed owner configuration builder used only during this Configure call; register this owner's concrete children.
END_VAR
VAR
    TestConfig : ST_TestCaseConfig;
END_VAR
Builder.Initialize(Mode := E_OrchestrationMode.Serial,
    TestCases := FTestCases);
FSignedRelations.Initialize(Parent := THIS^,
    TestName := 'SignedRelations',
    Config := TestConfig);
Builder.Register(TestCase := FSignedRelations);
FUnsignedRelations.Initialize(Parent := THIS^,
    TestName := 'UnsignedRelations',
    Config := TestConfig);
Builder.Register(TestCase := FUnsignedRelations);
FBitEquality.Initialize(Parent := THIS^,
    TestName := 'BitEquality',
    Config := TestConfig);
Builder.Register(TestCase := FBitEquality);
FBooleanComparisons.Initialize(Parent := THIS^,
    TestName := 'BooleanComparisons',
    Config := TestConfig);
Builder.Register(TestCase := FBooleanComparisons);
FCharacterEquality.Initialize(Parent := THIS^,
    TestName := 'CharacterEquality',
    Config := TestConfig);
Builder.Register(TestCase := FCharacterEquality);
FSignedRanges.Initialize(Parent := THIS^,
    TestName := 'SignedRanges',
    Config := TestConfig);
Builder.Register(TestCase := FSignedRanges);
FUnsignedRanges.Initialize(Parent := THIS^,
    TestName := 'UnsignedRanges',
    Config := TestConfig);
Builder.Register(TestCase := FUnsignedRanges);
FDurationComparisons.Initialize(Parent := THIS^,
    TestName := 'DurationComparisons',
    Config := TestConfig);
Builder.Register(TestCase := FDurationComparisons);
FDateNormalization.Initialize(Parent := THIS^,
    TestName := 'DateNormalization',
    Config := TestConfig);
Builder.Register(TestCase := FDateNormalization);
FTODDomain.Initialize(Parent := THIS^,
    TestName := 'TODDomain',
    Config := TestConfig);
Builder.Register(TestCase := FTODDomain);
FLTODDomain.Initialize(Parent := THIS^,
    TestName := 'LTODDomain',
    Config := TestConfig);
Builder.Register(TestCase := FLTODDomain);
FScalarDiagnostics.Initialize(Parent := THIS^,
    TestName := 'ScalarDiagnostics',
    Config := TestConfig);
Builder.Register(TestCase := FScalarDiagnostics);
END_METHOD

{region 'Documentation'}
(*!
<summary>Returns a registered scenario using its original array index.</summary>
*)
{endregion}
METHOD PUBLIC GetTestCase : I_TestCase //! Typed child interface at the original array index; zero when no entry is available.
VAR_INPUT
    Index : DINT; //! Original occupied child-array index, rather than an ordinal position.
END_VAR
GetTestCase := 0;
IF (ChildCount = 0) OR (Index < ChildArrayLowerBound)
    OR (DINT_TO_LINT(Index) >= DINT_TO_LINT(ChildArrayLowerBound) + UINT_TO_LINT(ChildCount)) THEN
    RETURN;
END_IF;
GetTestCase := FTestCases[Index];
END_METHOD

{region 'Documentation'}
(*!
<summary>Calls each owned scenario once per initialized Suite cycle.</summary>
*)
{endregion}
METHOD PROTECTED ProcessTestCases
FSignedRelations();
FUnsignedRelations();
FBitEquality();
FBooleanComparisons();
FCharacterEquality();
FSignedRanges();
FUnsignedRanges();
FDurationComparisons();
FDateNormalization();
FTODDomain();
FLTODDomain();
FScalarDiagnostics();
END_METHOD

END_FUNCTION_BLOCK

// ---- SelfTests/TestCases/TestSuite_AssertionComparisons/Test_AssertionSignedRelations.TcPOU
{region 'Documentation'}
(*!
<summary>Checks six native LINT comparison relations and full-width boundaries.</summary>
<description>
Each named row has explicit expected results, not a second comparison algorithm.
One disabled subject call consumes Reset before one enabled comparison call.
Outer checking Assertions latch every row before inputs advance; intentional
subject failures remain in a Test-Case-owned Event Buffer, cleared between rows.
Only the checking Assertions contribute to the outer result.
</description>
*)
{endregion}
FUNCTION_BLOCK Test_AssertionSignedRelations EXTENDS TestCaseBase
VAR
    FEqualSubject : AssertEqual_LInt;
    FNotEqualSubject : AssertNotEqual_LInt;
    FLessThanSubject : AssertLessThan_LInt;
    FLessEqualSubject : AssertLessEqual_LInt;
    FGreaterThanSubject : AssertGreaterThan_LInt;
    FGreaterEqualSubject : AssertGreaterEqual_LInt;
    FActual : LINT;
    FReference : LINT;
    FExpectedEqualResult : E_Result;
    FExpectedNotEqualResult : E_Result;
    FExpectedLessThanResult : E_Result;
    FExpectedLessEqualResult : E_Result;
    FExpectedGreaterThanResult : E_Result;
    FExpectedGreaterEqualResult : E_Result;
    FCapture : EventBuffer;
    FEvents : ARRAY[1..CaptureLength] OF ST_Event;
    FCaptureFifo : ST_FifoStatus;
    FCaptureStatus : ST_EventBufferStatus;
    FRow : UINT;
    FRowPrepared : BOOL;
    FObservationReady : BOOL;
    FChecked : BOOL;
    FSetupValid : BOOL;
END_VAR
VAR
    FEqualResult : AssertTrue;
    FEqualResultMatches : BOOL;
    FNotEqualResult : AssertTrue;
    FNotEqualResultMatches : BOOL;
    FLessThanResult : AssertTrue;
    FLessThanResultMatches : BOOL;
    FLessEqualResult : AssertTrue;
    FLessEqualResultMatches : BOOL;
    FGreaterThanResult : AssertTrue;
    FGreaterThanResultMatches : BOOL;
    FGreaterEqualResult : AssertTrue;
    FGreaterEqualResultMatches : BOOL;
    FCaptureIntegrity : AssertTrue;
    FCaptureIntegrityMatches : BOOL;
END_VAR
VAR CONSTANT
    CaptureLength : UINT := 8;
    ExpectedFindingCount : UDINT := 3;
    BelowZero : UINT := 1;
    EqualZero : UINT := 2;
    AboveZero : UINT := 3;
    MinimumBelowMaximum : UINT := 4;
    MaximumAboveMinimum : UINT := 5;
    MinimumEqual : UINT := 6;
    MaximumEqual : UINT := 7;
    LastRow : UINT := MaximumEqual;
    LowestValue : LINT := LINT#-9223372036854775808;
    HighestValue : LINT := LINT#9223372036854775807;
END_VAR

SUPER^();

{region 'Documentation'}
(*!
<summary>Collects only outer checking Assertions, never intentional subject findings.</summary>
*)
{endregion}
METHOD PROTECTED AggregateResults
VAR_INPUT
    Aggregator : I_ResultAggregator; //! Borrowed result sink owned by the outer Test Case; add this test's checking Assertions without resetting or retaining the sink.
END_VAR
Aggregator.AddProvider(Provider := FEqualResult);
Aggregator.AddProvider(Provider := FNotEqualResult);
Aggregator.AddProvider(Provider := FLessThanResult);
Aggregator.AddProvider(Provider := FLessEqualResult);
Aggregator.AddProvider(Provider := FGreaterThanResult);
Aggregator.AddProvider(Provider := FGreaterEqualResult);
Aggregator.AddProvider(Provider := FCaptureIntegrity);
END_METHOD

{region 'Documentation'}
(*!
<summary>Calls each real comparison once with the selected typed row inputs.</summary>
*)
{endregion}
METHOD PRIVATE CallSubjects
VAR_INPUT
    Enable : BOOL; //! Observation-enable input forwarded to the controlled Assertion subjects for this call.
END_VAR
FEqualSubject(Enable := Enable,
    State := E_State.Running,
    IN := FActual,
    Expected := FReference);
FNotEqualSubject(Enable := Enable,
    State := E_State.Running,
    IN := FActual,
    Expected := FReference);
FLessThanSubject(Enable := Enable,
    State := E_State.Running,
    IN := FActual,
    Maximum := FReference);
FLessEqualSubject(Enable := Enable,
    State := E_State.Running,
    IN := FActual,
    Maximum := FReference);
FGreaterThanSubject(Enable := Enable,
    State := E_State.Running,
    IN := FActual,
    Minimum := FReference);
FGreaterEqualSubject(Enable := Enable,
    State := E_State.Running,
    IN := FActual,
    Minimum := FReference);
END_METHOD

{region 'Documentation'}
(*!
<summary>Preserves base validation and rejects incomplete subject or checking-Assertion setup.</summary>
*)
{endregion}
METHOD PROTECTED CheckInitialization : BOOL //! TRUE when the inherited initialization check and this concrete fixture check both accept the setup.
CheckInitialization := SUPER^.CheckInitialization();
IF NOT CheckInitialization THEN
    RETURN;
END_IF;

CheckInitialization := FSetupValid
    AND FEqualResult.IsInitialized
    AND FNotEqualResult.IsInitialized
    AND FLessThanResult.IsInitialized
    AND FLessEqualResult.IsInitialized
    AND FGreaterThanResult.IsInitialized
    AND FGreaterEqualResult.IsInitialized
    AND FCaptureIntegrity.IsInitialized;
IF NOT CheckInitialization THEN
    EventPublisher.PublishEvent(Event := CreateFrameworkEvent(Name := Name,
        ResourceName := '',
        State := State,
        Severity := E_EventSeverity.Error,
        Message := 'Comparison selftest setup failed.'));
END_IF;
END_METHOD

{region 'Documentation'}
(*!
<summary>Compares observed results with the literal row expectations and checks local event loss/count.</summary>
*)
{endregion}
METHOD PRIVATE CheckResults
FEqualResultMatches := FEqualSubject.Result = FExpectedEqualResult;
FNotEqualResultMatches := FNotEqualSubject.Result = FExpectedNotEqualResult;
FLessThanResultMatches := FLessThanSubject.Result = FExpectedLessThanResult;
FLessEqualResultMatches := FLessEqualSubject.Result = FExpectedLessEqualResult;
FGreaterThanResultMatches := FGreaterThanSubject.Result = FExpectedGreaterThanResult;
FGreaterEqualResultMatches := FGreaterEqualSubject.Result = FExpectedGreaterEqualResult;
FCaptureIntegrityMatches := (FCaptureStatus.SequenceId = ExpectedFindingCount)
    AND (FCaptureStatus.LostEventCount = 0);
END_METHOD

{region 'Documentation'}
(*!
<summary>Initializes the local capture, checking Assertions and publisher-bound real comparisons.</summary>
*)
{endregion}
METHOD PROTECTED Configure
VAR
    Initialized : BOOL;
END_VAR
FPreparationStateCount := 0;
FTestStateCount := 1;
FEqualResult.Initialize(Parent := THIS^,
    AssertionName := 'EqualResult');
FNotEqualResult.Initialize(Parent := THIS^,
    AssertionName := 'NotEqualResult');
FLessThanResult.Initialize(Parent := THIS^,
    AssertionName := 'LessThanResult');
FLessEqualResult.Initialize(Parent := THIS^,
    AssertionName := 'LessEqualResult');
FGreaterThanResult.Initialize(Parent := THIS^,
    AssertionName := 'GreaterThanResult');
FGreaterEqualResult.Initialize(Parent := THIS^,
    AssertionName := 'GreaterEqualResult');
FCaptureIntegrity.Initialize(Parent := THIS^,
    AssertionName := 'CaptureIntegrity');
FSetupValid := FCapture.Initialize(Buffer := FEvents,
    FifoControl := FCaptureFifo,
    Status := FCaptureStatus);
FEqualSubject.BindPublisher(Publisher := FCapture);
Initialized := FEqualSubject.Initialize(Parent := THIS^,
    AssertionName := 'EqualSubject');
FSetupValid := FSetupValid AND Initialized;
FNotEqualSubject.BindPublisher(Publisher := FCapture);
Initialized := FNotEqualSubject.Initialize(Parent := THIS^,
    AssertionName := 'NotEqualSubject');
FSetupValid := FSetupValid AND Initialized;
FLessThanSubject.BindPublisher(Publisher := FCapture);
Initialized := FLessThanSubject.Initialize(Parent := THIS^,
    AssertionName := 'LessThanSubject');
FSetupValid := FSetupValid AND Initialized;
FLessEqualSubject.BindPublisher(Publisher := FCapture);
Initialized := FLessEqualSubject.Initialize(Parent := THIS^,
    AssertionName := 'LessEqualSubject');
FSetupValid := FSetupValid AND Initialized;
FGreaterThanSubject.BindPublisher(Publisher := FCapture);
Initialized := FGreaterThanSubject.Initialize(Parent := THIS^,
    AssertionName := 'GreaterThanSubject');
FSetupValid := FSetupValid AND Initialized;
FGreaterEqualSubject.BindPublisher(Publisher := FCapture);
Initialized := FGreaterEqualSubject.Initialize(Parent := THIS^,
    AssertionName := 'GreaterEqualSubject');
FSetupValid := FSetupValid AND Initialized;
END_METHOD

{region 'Documentation'}
(*!
<summary>Completes abort without asynchronous resources.</summary>
*)
{endregion}
METHOD PROTECTED ProcessAbort
VAR_INPUT
    Enable : BOOL; //! Phase permission supplied by the owning Test Case; FALSE does not authorize progression, while observation may continue.
END_VAR
IF Enable THEN
    CompleteAbort();
END_IF;
END_METHOD

{region 'Documentation'}
(*!
<summary>Latches checked observations before the next script step may proceed.</summary>
*)
{endregion}
METHOD PROTECTED ProcessAssertions
VAR_INPUT
    Enable : BOOL; //! Phase permission supplied by the owning Test Case; FALSE does not authorize progression, while observation may continue.
END_VAR
VAR
    Evaluate : BOOL;
END_VAR
Evaluate := Enable AND FObservationReady;
FEqualResult(Enable := Evaluate,
    State := State,
    IN := FEqualResultMatches);
FNotEqualResult(Enable := Evaluate,
    State := State,
    IN := FNotEqualResultMatches);
FLessThanResult(Enable := Evaluate,
    State := State,
    IN := FLessThanResultMatches);
FLessEqualResult(Enable := Evaluate,
    State := State,
    IN := FLessEqualResultMatches);
FGreaterThanResult(Enable := Evaluate,
    State := State,
    IN := FGreaterThanResultMatches);
FGreaterEqualResult(Enable := Evaluate,
    State := State,
    IN := FGreaterEqualResultMatches);
FCaptureIntegrity(Enable := Evaluate,
    State := State,
    IN := FCaptureIntegrityMatches);
IF Evaluate THEN
    FChecked := TRUE;
END_IF;
END_METHOD

{region 'Documentation'}
(*!
<summary>No Preparation phase is required.</summary>
*)
{endregion}
METHOD PROTECTED ProcessPreparations
VAR_INPUT
    // SA0033: Required hook; this test has no Preparation phase.
    {attribute 'analysis' := '-33'}
    Enable : BOOL; //! Phase permission supplied by the owning Test Case; FALSE does not authorize progression, while observation may continue.
END_VAR
END_METHOD

{region 'Documentation'}
(*!
<summary>Restarts the script and resets the checking Assertions.</summary>
*)
{endregion}
METHOD PROTECTED ProcessReset
FRow := BelowZero;
FRowPrepared := FALSE;
FChecked := FALSE;
FObservationReady := FALSE;
FEqualResult.Reset();
FEqualResultMatches := TRUE;
FNotEqualResult.Reset();
FNotEqualResultMatches := TRUE;
FLessThanResult.Reset();
FLessThanResultMatches := TRUE;
FLessEqualResult.Reset();
FLessEqualResultMatches := TRUE;
FGreaterThanResult.Reset();
FGreaterThanResultMatches := TRUE;
FGreaterEqualResult.Reset();
FGreaterEqualResultMatches := TRUE;
FCaptureIntegrity.Reset();
FCaptureIntegrityMatches := TRUE;
CompleteReset();
END_METHOD

{region 'Documentation'}
(*!
<summary>Advances one bounded script step per active PLC cycle.</summary>
*)
{endregion}
METHOD PROTECTED ProcessTests
VAR_INPUT
    Enable : BOOL; //! Phase permission supplied by the owning Test Case; FALSE does not authorize progression, while observation may continue.
END_VAR
IF NOT Enable THEN
    RETURN;
END_IF;

IF FChecked THEN
    FChecked := FALSE;
    FObservationReady := FALSE;
    IF FRow = LastRow THEN
        CompleteTests();
        RETURN;
    END_IF;
    FRow := FRow + 1;
    FRowPrepared := FALSE;
END_IF;

IF NOT FRowPrepared THEN
    SelectRow();
    FCapture.Reset();
    ResetSubjects();
    CallSubjects(Enable := FALSE);
    FRowPrepared := TRUE;
ELSE
    CallSubjects(Enable := TRUE);
    CheckResults();
    FObservationReady := TRUE;
END_IF;
END_METHOD

{region 'Documentation'}
(*!
<summary>Requests a fresh result epoch for every comparison; CallSubjects consumes it.</summary>
*)
{endregion}
METHOD PRIVATE ResetSubjects
FEqualSubject.Reset();
FNotEqualSubject.Reset();
FLessThanSubject.Reset();
FLessEqualSubject.Reset();
FGreaterThanSubject.Reset();
FGreaterEqualSubject.Reset();
END_METHOD

